// TwinCAT 3 PLC project Syn_Visu_Test
// ProgramVersion: 3.1.4026.28
// libraries:
//   Tc2_Standard, * (Beckhoff Automation GmbH)
//   Tc2_System, * (Beckhoff Automation GmbH)
//   SynConfig,newest,Syntegon Group
//   SynVisu,newest,Syntegon Group
//   TcUnit,newest,www.tcunit.org
// project tree:
//   / PlcTask.TcTTO
//   POUs/ P_TestRun.TcPOU
//   POUs/Tests/ _FB_TestBodyComponent.TcPOU, _FB_TestComponent.TcPOU, _FB_TestConfigBodyComponent.TcPOU, _FB_TestConfigComponent.TcPOU, _FB_TestConfigMachine.TcPOU, _FB_TestConfigRobot.TcPOU, _FB_TestConfigStaging.TcPOU, _FB_TestConfigTopology.TcPOU, _FB_TestConveyor.TcPOU, _FB_TestMachine.TcPOU, _FB_TestProductRegister.TcPOU, _FB_TestRobot.TcPOU, _FB_TestXtsTrack.TcPOU, _FC_TestConfigStage.TcPOU
// (motion and I/O tree: see PLC project syn_visu)
// real-time tasks:
//   TASK PlcTask: cycle T#10ms, priority 20, ADS port 350
//   TASK TestTask: cycle T#10ms, priority 21, ADS port 351

CONFIGURATION Syn_Visu_Test
    RESOURCE PLC ON TwinCAT3
        TASK PlcTask(INTERVAL := T#10ms, PRIORITY := 21);
        PROGRAM P_TestRun WITH PlcTask : P_TestRun;
    END_RESOURCE
END_CONFIGURATION

// ---- POUs/P_TestRun.TcPOU
(****************************************************************************************************<br>
© Syntegon Group.<br>
All rights reserved, also regarding any disposal, exploitation, reproduction, editing, distribution,<br>
as well as in the event of applications for industrial property rights.<br>
*****************************************************************************************************<br>
DESCRIPTION:<br>
Runs the TcUnit unit tests of the libraries Syn_Visu and Syn_Config (the installed SynVisu and SynConfig, newest<br>
versions) once after the start: every suite in POUs/Tests (_FB_TestConfig... for Syn_Config). TcUnit writes the<br>
results to the error list (ADS log) and, through TcUnit-Runner, to an xUnit file. Tests use only the libraries'<br>
public methods and their contract structures, written as the gateway writes them.<br>
****************************************************************************************************)
PROGRAM P_TestRun
VAR
	fb_TestComponent					: _FB_TestComponent;
	fb_TestConveyor						: _FB_TestConveyor;
	fb_TestProductRegister				: _FB_TestProductRegister;
	fb_TestRobot						: _FB_TestRobot;
	fb_TestXtsTrack						: _FB_TestXtsTrack;
	fb_TestBodyComponent				: _FB_TestBodyComponent;
	fb_TestMachine						: _FB_TestMachine;
	fb_TestConfigComponent				: _FB_TestConfigComponent;
	fb_TestConfigStaging				: _FB_TestConfigStaging;
	fb_TestConfigRobot					: _FB_TestConfigRobot;
	fb_TestConfigBodyComponent			: _FB_TestConfigBodyComponent;
	fb_TestConfigMachine				: _FB_TestConfigMachine;
	fb_TestConfigTopology				: _FB_TestConfigTopology;
END_VAR

TcUnit.RUN();

END_PROGRAM

// ---- POUs/Tests/_FB_TestComponent.TcPOU
(****************************************************************************************************<br>
© Syntegon Group.<br>
All rights reserved, also regarding any disposal, exploitation, reproduction, editing, distribution,<br>
as well as in the event of applications for industrial property rights.<br>
*****************************************************************************************************<br>
DESCRIPTION:<br>
TcUnit test suite of _FB_VisuComponent: registration in the manifest (m_Register, m_Id), the symbol path<br>
taken from the instance path, and the library version reported to the gateway.<br>
*****************************************************************************************************<br>
VERSION         ¦ DATE       ¦ NAME      ¦ CHANGE<br>
Syn_Visu 9.4.0  ¦ 2026-11-09 ¦ J.Willner ¦ Unit tests<br>
Syn_Visu 10.0.0 ¦ 2026-11-14 ¦ J.Willner ¦ _FC_VisuSymbolPath<br>
****************************************************************************************************)
FUNCTION_BLOCK _FB_TestComponent EXTENDS TcUnit.FB_TestSuite
VAR
	fb_PathConveyor						: _FB_VisuConveyor;	// declared here so that its instance path is known
END_VAR

m_RegisterAddsEntry();
m_RegisterIsIdempotent();
m_RegisterRejectsIdZero();
m_RegisterRejectsUsedId();
m_RegisterRejectsFullManifest();
m_RegisterSymbolPath();
m_SymbolPathFromInstancePath();
m_VersionMatchesConstant();

(****************************************************************************************************<br>
© Syntegon Group.<br>
All rights reserved, also regarding any disposal, exploitation, reproduction, editing, distribution,<br>
as well as in the event of applications for industrial property rights.<br>
*****************************************************************************************************<br>
DESCRIPTION:<br>
A new component gets a manifest entry with its id, type and name; the config version goes up by one and the<br>
manifest reports the running library's protocol and library version.<br>
****************************************************************************************************)
METHOD PRIVATE m_RegisterAddsEntry
VAR_INST
	fb_TempConveyor						: _FB_VisuConveyor;
	TempManifest						: ST_VisuManifest;
	b_TempDone							: BOOL;	// the test ran
END_VAR
TEST('RegisterAddsEntry');
IF b_TempDone THEN
	RETURN;
END_IF
b_TempDone := TRUE;

TempManifest.nProtocolVersion := 0;
AssertTrue(Condition := fb_TempConveyor.m_Register(vio_Manifest := TempManifest, vi_udn_Id := 1, vi_str_Name := 'Infeed'),
	Message := 'm_Register accepts a new id');
AssertEquals_UINT(Expected := 1, Actual := TempManifest.nCount, Message := 'one manifest entry');
AssertEquals_UDINT(Expected := 1, Actual := TempManifest.aEntries[0].nId, Message := 'entry id');
AssertTrue(Condition := TempManifest.aEntries[0].eType = E_VisuComponentType.CONVEYOR, Message := 'entry type CONVEYOR');
AssertEquals_STRING(Expected := 'Infeed', Actual := TempManifest.aEntries[0].sName, Message := 'entry name');
AssertEquals_UDINT(Expected := 2, Actual := TempManifest.nConfigVersion, Message := 'config version 1 -> 2');
AssertEquals_UINT(Expected := VISU_GlobalConst.VISU_un_PROTOCOL_VERSION, Actual := TempManifest.nProtocolVersion,
	Message := 'protocol version reported');
AssertEquals_STRING(Expected := VISU_GlobalConst.VISU_str_LIBRARY_VERSION, Actual := TempManifest.sLibraryVersion,
	Message := 'library version reported');
AssertEquals_UDINT(Expected := 1, Actual := fb_TempConveyor.m_Id(), Message := 'm_Id gives the registered id');

TEST_FINISHED();
END_METHOD

(****************************************************************************************************<br>
© Syntegon Group.<br>
All rights reserved, also regarding any disposal, exploitation, reproduction, editing, distribution,<br>
as well as in the event of applications for industrial property rights.<br>
*****************************************************************************************************<br>
DESCRIPTION:<br>
m_Register is called every cycle: registering again with the same values keeps the single entry and the<br>
config version.<br>
****************************************************************************************************)
METHOD PRIVATE m_RegisterIsIdempotent
VAR_INST
	fb_TempConveyor						: _FB_VisuConveyor;
	TempManifest						: ST_VisuManifest;
	b_TempDone							: BOOL;	// the test ran
END_VAR
TEST('RegisterIsIdempotent');
IF b_TempDone THEN
	RETURN;
END_IF
b_TempDone := TRUE;

fb_TempConveyor.m_Register(vio_Manifest := TempManifest, vi_udn_Id := 3, vi_str_Name := 'Outfeed');
AssertTrue(Condition := fb_TempConveyor.m_Register(vio_Manifest := TempManifest, vi_udn_Id := 3, vi_str_Name := 'Outfeed'),
	Message := 'the second m_Register with the same values succeeds');
AssertEquals_UINT(Expected := 1, Actual := TempManifest.nCount, Message := 'still one manifest entry');
AssertEquals_UDINT(Expected := 2, Actual := TempManifest.nConfigVersion, Message := 'config version unchanged by the second call');

TEST_FINISHED();
END_METHOD

(****************************************************************************************************<br>
© Syntegon Group.<br>
All rights reserved, also regarding any disposal, exploitation, reproduction, editing, distribution,<br>
as well as in the event of applications for industrial property rights.<br>
*****************************************************************************************************<br>
DESCRIPTION:<br>
A manifest holding VISU_un_MAX_MANIFEST_ENTRIES entries takes no further component.<br>
****************************************************************************************************)
METHOD PRIVATE m_RegisterRejectsFullManifest
VAR_INST
	fb_TempConveyor						: _FB_VisuConveyor;
	TempManifest						: ST_VisuManifest;
	b_TempDone							: BOOL;	// the test ran
END_VAR
TEST('RegisterRejectsFullManifest');
IF b_TempDone THEN
	RETURN;
END_IF
b_TempDone := TRUE;

(* Entries with id 0 never match a new id, so the manifest only counts as full. *)
TempManifest.nCount := VISU_GlobalConst_Param.VISU_un_MAX_MANIFEST_ENTRIES;
AssertFalse(Condition := fb_TempConveyor.m_Register(vio_Manifest := TempManifest, vi_udn_Id := 1, vi_str_Name := 'Infeed'),
	Message := 'full manifest refuses a new entry');
AssertEquals_UINT(Expected := VISU_GlobalConst_Param.VISU_un_MAX_MANIFEST_ENTRIES, Actual := TempManifest.nCount,
	Message := 'entry count unchanged');
AssertEquals_UDINT(Expected := 1, Actual := TempManifest.nConfigVersion, Message := 'config version unchanged');

TEST_FINISHED();
END_METHOD

(****************************************************************************************************<br>
© Syntegon Group.<br>
All rights reserved, also regarding any disposal, exploitation, reproduction, editing, distribution,<br>
as well as in the event of applications for industrial property rights.<br>
*****************************************************************************************************<br>
DESCRIPTION:<br>
Id 0 is refused without an entry, but the manifest still reports the running library's versions.<br>
****************************************************************************************************)
METHOD PRIVATE m_RegisterRejectsIdZero
VAR_INST
	fb_TempConveyor						: _FB_VisuConveyor;
	TempManifest						: ST_VisuManifest;
	b_TempDone							: BOOL;	// the test ran
END_VAR
TEST('RegisterRejectsIdZero');
IF b_TempDone THEN
	RETURN;
END_IF
b_TempDone := TRUE;

TempManifest.nProtocolVersion := 0;
AssertFalse(Condition := fb_TempConveyor.m_Register(vio_Manifest := TempManifest, vi_udn_Id := 0, vi_str_Name := 'Infeed'),
	Message := 'm_Register refuses id 0');
AssertEquals_UINT(Expected := 0, Actual := TempManifest.nCount, Message := 'no manifest entry');
AssertEquals_UDINT(Expected := 1, Actual := TempManifest.nConfigVersion, Message := 'config version unchanged');
AssertEquals_UDINT(Expected := 0, Actual := fb_TempConveyor.m_Id(), Message := 'm_Id stays 0');
AssertEquals_UINT(Expected := VISU_GlobalConst.VISU_un_PROTOCOL_VERSION, Actual := TempManifest.nProtocolVersion,
	Message := 'protocol version reported anyway');

TEST_FINISHED();
END_METHOD

(****************************************************************************************************<br>
© Syntegon Group.<br>
All rights reserved, also regarding any disposal, exploitation, reproduction, editing, distribution,<br>
as well as in the event of applications for industrial property rights.<br>
*****************************************************************************************************<br>
DESCRIPTION:<br>
An id already used by a different entry (other type or other name) is refused; the first entry stays.<br>
****************************************************************************************************)
METHOD PRIVATE m_RegisterRejectsUsedId
VAR_INST
	fb_TempConveyor						: _FB_VisuConveyor;
	fb_TempOtherConveyor				: _FB_VisuConveyor;
	fb_TempDelta						: _FB_VisuDelta;
	TempManifest						: ST_VisuManifest;
	b_TempDone							: BOOL;	// the test ran
END_VAR
TEST('RegisterRejectsUsedId');
IF b_TempDone THEN
	RETURN;
END_IF
b_TempDone := TRUE;

fb_TempConveyor.m_Register(vio_Manifest := TempManifest, vi_udn_Id := 5, vi_str_Name := 'Infeed');
AssertFalse(Condition := fb_TempDelta.m_Register(vio_Manifest := TempManifest, vi_udn_Id := 5, vi_str_Name := 'Infeed'),
	Message := 'same id, other type: refused');
AssertFalse(Condition := fb_TempOtherConveyor.m_Register(vio_Manifest := TempManifest, vi_udn_Id := 5, vi_str_Name := 'Other'),
	Message := 'same id, other name: refused');
AssertEquals_UINT(Expected := 1, Actual := TempManifest.nCount, Message := 'still one manifest entry');
AssertEquals_UDINT(Expected := 0, Actual := fb_TempDelta.m_Id(), Message := 'refused component keeps m_Id 0');
AssertEquals_UDINT(Expected := 5, Actual := fb_TempConveyor.m_Id(), Message := 'first component keeps its id');

TEST_FINISHED();
END_METHOD

(****************************************************************************************************<br>
© Syntegon Group.<br>
All rights reserved, also regarding any disposal, exploitation, reproduction, editing, distribution,<br>
as well as in the event of applications for industrial property rights.<br>
*****************************************************************************************************<br>
DESCRIPTION:<br>
The manifest entry's symbol path is the instance path without TwinCAT project and PLC project, plus<br>
'.vo_Visu': the path the gateway reads over ADS.<br>
****************************************************************************************************)
METHOD PRIVATE m_RegisterSymbolPath
VAR_INST
	TempManifest						: ST_VisuManifest;
	b_TempDone							: BOOL;	// the test ran
END_VAR
TEST('RegisterSymbolPath');
IF b_TempDone THEN
	RETURN;
END_IF
b_TempDone := TRUE;

fb_PathConveyor.m_Register(vio_Manifest := TempManifest, vi_udn_Id := 1, vi_str_Name := 'Path');
AssertEquals_STRING(Expected := 'P_TestRun.fb_TestComponent.fb_PathConveyor.vo_Visu', Actual := TempManifest.aEntries[0].sPath,
	Message := 'symbol path of vo_Visu without TwinCAT and PLC project');

TEST_FINISHED();
END_METHOD

(****************************************************************************************************<br>
© Syntegon Group.<br>
All rights reserved, also regarding any disposal, exploitation, reproduction, editing, distribution,<br>
as well as in the event of applications for industrial property rights.<br>
*****************************************************************************************************<br>
DESCRIPTION:<br>
_FC_VisuSymbolPath, the rule both manifests use: the instance path without TwinCAT project and PLC project,<br>
plus the contract structure; a path with fewer segments is kept whole.<br>
****************************************************************************************************)
METHOD PRIVATE m_SymbolPathFromInstancePath
VAR_INST
	b_TempDone							: BOOL;	// the test ran
END_VAR
TEST('SymbolPathFromInstancePath');
IF b_TempDone THEN
	RETURN;
END_IF
b_TempDone := TRUE;

AssertEquals_STRING(Expected := 'P_VisuDemoDelta.fb_Infeed1.vo_Visu',
	Actual := _FC_VisuSymbolPath(vio_str_InstancePath := 'RPP_Visu.Syn_Visu_Demo.P_VisuDemoDelta.fb_Infeed1',
		vi_str_Member := '.vo_Visu'), Message := 'TwinCAT and PLC project left out');
AssertEquals_STRING(Expected := 'P_A.fb_B.vo_Config',
	Actual := _FC_VisuSymbolPath(vio_str_InstancePath := 'Tc.Plc.P_A.fb_B', vi_str_Member := '.vo_Config'),
	Message := 'another contract structure');
AssertEquals_STRING(Expected := 'MAIN.fb_A.vo_Visu',
	Actual := _FC_VisuSymbolPath(vio_str_InstancePath := 'MAIN.fb_A', vi_str_Member := '.vo_Visu'),
	Message := 'fewer segments: kept whole');

TEST_FINISHED();
END_METHOD

(****************************************************************************************************<br>
© Syntegon Group.<br>
All rights reserved, also regarding any disposal, exploitation, reproduction, editing, distribution,<br>
as well as in the event of applications for industrial property rights.<br>
*****************************************************************************************************<br>
DESCRIPTION:<br>
_FC_GetVersionSynVisu and VISU_str_LIBRARY_VERSION name the same version: both are bumped together.<br>
****************************************************************************************************)
METHOD PRIVATE m_VersionMatchesConstant
VAR_INST
	b_TempDone							: BOOL;	// the test ran
END_VAR
VAR
	str_TempVersion						: STRING(31);	// major.minor.revision from _FC_GetVersionSynVisu
END_VAR
TEST('VersionMatchesConstant');
IF b_TempDone THEN
	RETURN;
END_IF
b_TempDone := TRUE;

str_TempVersion := CONCAT(UINT_TO_STRING(_FC_GetVersionSynVisu(vi_n_VersionElement := 1)), '.');
str_TempVersion := CONCAT(str_TempVersion, UINT_TO_STRING(_FC_GetVersionSynVisu(vi_n_VersionElement := 2)));
str_TempVersion := CONCAT(str_TempVersion, '.');
str_TempVersion := CONCAT(str_TempVersion, UINT_TO_STRING(_FC_GetVersionSynVisu(vi_n_VersionElement := 3)));
AssertEquals_STRING(Expected := VISU_GlobalConst.VISU_str_LIBRARY_VERSION, Actual := str_TempVersion,
	Message := '_FC_GetVersionSynVisu matches VISU_str_LIBRARY_VERSION');
AssertEquals_UINT(Expected := 16#FFFF, Actual := _FC_GetVersionSynVisu(vi_n_VersionElement := 4),
	Message := 'unknown version element gives 16#FFFF');

TEST_FINISHED();
END_METHOD

END_FUNCTION_BLOCK

// ---- POUs/Tests/_FB_TestConveyor.TcPOU
(****************************************************************************************************<br>
© Syntegon Group.<br>
All rights reserved, also regarding any disposal, exploitation, reproduction, editing, distribution,<br>
as well as in the event of applications for industrial property rights.<br>
*****************************************************************************************************<br>
DESCRIPTION:<br>
TcUnit test suite of _FB_VisuConveyor's config and belt position: the config version only changes when a<br>
value does, product types, the body flag, the unwrapping of a modulo belt position and the conversion between<br>
the MCS and the conveyor's coordinate system.<br>
*****************************************************************************************************<br>
VERSION         ¦ DATE       ¦ NAME      ¦ CHANGE<br>
Syn_Visu 9.4.0  ¦ 2026-11-09 ¦ J.Willner ¦ Unit tests<br>
Syn_Visu 10.0.0 ¦ 2026-11-14 ¦ J.Willner ¦ m_SetPose; m_BeltToMcs and m_McsToBelt<br>
****************************************************************************************************)
FUNCTION_BLOCK _FB_TestConveyor EXTENDS TcUnit.FB_TestSuite

m_ConfigureChangesVersionOnce();
m_SetProductTypeAddsAndUpdates();
m_SetProductTypeRejectsFullList();
m_SetBodyVisible();
m_SetModuloBeltPosition();
m_BeltAndMcsConvert();

(****************************************************************************************************<br>
© Syntegon Group.<br>
All rights reserved, also regarding any disposal, exploitation, reproduction, editing, distribution,<br>
as well as in the event of applications for industrial property rights.<br>
*****************************************************************************************************<br>
DESCRIPTION:<br>
m_BeltToMcs places a pose of the conveyor's coordinate system in the MCS as the visualisation does (the pose's<br>
rotation turns the origin shift and the position, fRz adds up), and m_McsToBelt is its inverse, also on a<br>
tilted conveyor.<br>
****************************************************************************************************)
METHOD PRIVATE m_BeltAndMcsConvert
VAR_INST
	fb_TempConveyor						: _FB_VisuConveyor;
	b_TempDone							: BOOL;	// the test ran
END_VAR
VAR
	TempPose							: ST_VisuPose;	// of the conveyor
	TempBelt							: ST_VisuPlanarPose;	// conveyor coordinate system
	TempMcs								: ST_VisuPlanarPose;
END_VAR
TEST('BeltAndMcsConvert');
IF b_TempDone THEN
	RETURN;
END_IF
b_TempDone := TRUE;


(****************************************************************************************************
A CONVEYOR TURNED BY 90 DEGREES
****************************************************************************************************)
TempPose.fX := 1000;
TempPose.fY := 500;
TempPose.fZ := 800;
TempPose.fRz := 90;
fb_TempConveyor.m_SetPose(vi_Pose := TempPose);
fb_TempConveyor.m_SetOriginShift(vi_lr_X := 100, vi_lr_Y := 0, vi_lr_Z := 0);

(* Its coordinate system lies 100 mm along the belt, i.e. along the MCS +Y. *)
TempMcs := fb_TempConveyor.m_BeltToMcs(vi_Pose := TempBelt);
AssertEquals_LREAL(Expected := 1000, Actual := TempMcs.fX, Delta := 0.001, Message := 'origin X');
AssertEquals_LREAL(Expected := 600, Actual := TempMcs.fY, Delta := 0.001, Message := 'origin Y');
AssertEquals_LREAL(Expected := 800, Actual := TempMcs.fZ, Delta := 0.001, Message := 'origin Z');
AssertEquals_LREAL(Expected := 90, Actual := TempMcs.fRz, Delta := 0.001, Message := 'origin Rz');

TempBelt.fX := 50;
TempBelt.fY := 20;
TempBelt.fZ := 10;
TempBelt.fRz := 15;
TempMcs := fb_TempConveyor.m_BeltToMcs(vi_Pose := TempBelt);
AssertEquals_LREAL(Expected := 980, Actual := TempMcs.fX, Delta := 0.001, Message := 'belt Y runs along MCS -X');
AssertEquals_LREAL(Expected := 650, Actual := TempMcs.fY, Delta := 0.001, Message := 'belt X runs along MCS +Y');
AssertEquals_LREAL(Expected := 810, Actual := TempMcs.fZ, Delta := 0.001, Message := 'Z');
AssertEquals_LREAL(Expected := 105, Actual := TempMcs.fRz, Delta := 0.001, Message := 'Rz adds up');

TempBelt := fb_TempConveyor.m_McsToBelt(vi_Pose := TempMcs);
AssertEquals_LREAL(Expected := 50, Actual := TempBelt.fX, Delta := 0.001, Message := 'back: X');
AssertEquals_LREAL(Expected := 20, Actual := TempBelt.fY, Delta := 0.001, Message := 'back: Y');
AssertEquals_LREAL(Expected := 10, Actual := TempBelt.fZ, Delta := 0.001, Message := 'back: Z');
AssertEquals_LREAL(Expected := 15, Actual := TempBelt.fRz, Delta := 0.001, Message := 'back: Rz');


(****************************************************************************************************
A TILTED CONVEYOR: THERE AND BACK
****************************************************************************************************)
TempPose.fRx := 5;
TempPose.fRy := -3;
TempPose.fRz := 30;
fb_TempConveyor.m_SetPose(vi_Pose := TempPose);
fb_TempConveyor.m_SetOriginShift(vi_lr_X := 100, vi_lr_Y := -40, vi_lr_Z := 25);
TempBelt.fX := 321;
TempBelt.fY := -45;
TempBelt.fZ := 12;
TempBelt.fRz := 7;
TempBelt := fb_TempConveyor.m_McsToBelt(vi_Pose := fb_TempConveyor.m_BeltToMcs(vi_Pose := TempBelt));
AssertEquals_LREAL(Expected := 321, Actual := TempBelt.fX, Delta := 0.001, Message := 'tilted: X');
AssertEquals_LREAL(Expected := -45, Actual := TempBelt.fY, Delta := 0.001, Message := 'tilted: Y');
AssertEquals_LREAL(Expected := 12, Actual := TempBelt.fZ, Delta := 0.001, Message := 'tilted: Z');
AssertEquals_LREAL(Expected := 7, Actual := TempBelt.fRz, Delta := 0.001, Message := 'tilted: Rz');

TEST_FINISHED();
END_METHOD

(****************************************************************************************************<br>
© Syntegon Group.<br>
All rights reserved, also regarding any disposal, exploitation, reproduction, editing, distribution,<br>
as well as in the event of applications for industrial property rights.<br>
*****************************************************************************************************<br>
DESCRIPTION:<br>
m_SetPose and m_Configure may be called every cycle: only a changed value raises the manifest's config version.<br>
****************************************************************************************************)
METHOD PRIVATE m_ConfigureChangesVersionOnce
VAR_INST
	fb_TempConveyor						: _FB_VisuConveyor;
	TempManifest						: ST_VisuManifest;
	TempPose							: ST_VisuPose;
	b_TempDone							: BOOL;	// the test ran
END_VAR
VAR
	udn_TempVersion						: UDINT;	// [-] config version after m_Register
END_VAR
TEST('ConfigureChangesVersionOnce');
IF b_TempDone THEN
	RETURN;
END_IF
b_TempDone := TRUE;

fb_TempConveyor.m_Register(vio_Manifest := TempManifest, vi_udn_Id := 1, vi_str_Name := 'Infeed');
udn_TempVersion := TempManifest.nConfigVersion;
TempPose.fX := 100;
AssertTrue(Condition := fb_TempConveyor.m_SetPose(vi_Pose := TempPose), Message := 'first m_SetPose changes the config');
AssertTrue(Condition := fb_TempConveyor.m_Configure(vi_lr_Length := 3000, vi_lr_Width := 400),
	Message := 'first m_Configure changes the config');
AssertEquals_UDINT(Expected := udn_TempVersion + 2, Actual := TempManifest.nConfigVersion,
	Message := 'config version raised once by each');
AssertFalse(Condition := fb_TempConveyor.m_SetPose(vi_Pose := TempPose), Message := 'same pose: no change');
AssertFalse(Condition := fb_TempConveyor.m_Configure(vi_lr_Length := 3000, vi_lr_Width := 400),
	Message := 'same values: no change');
AssertEquals_UDINT(Expected := udn_TempVersion + 2, Actual := TempManifest.nConfigVersion, Message := 'config version unchanged');
AssertTrue(Condition := fb_TempConveyor.m_Configure(vi_lr_Length := 3500, vi_lr_Width := 400),
	Message := 'new length changes the config');
AssertEquals_UDINT(Expected := udn_TempVersion + 3, Actual := TempManifest.nConfigVersion, Message := 'config version raised again');
AssertEquals_LREAL(Expected := 3500, Actual := fb_TempConveyor.vo_Visu.stConfig.fLength, Delta := 0.001,
	Message := 'length taken over');
AssertEquals_LREAL(Expected := 100, Actual := fb_TempConveyor.vo_Visu.stConfig.stPose.fX, Delta := 0.001,
	Message := 'pose kept by m_Configure');

TEST_FINISHED();
END_METHOD

(****************************************************************************************************<br>
© Syntegon Group.<br>
All rights reserved, also regarding any disposal, exploitation, reproduction, editing, distribution,<br>
as well as in the event of applications for industrial property rights.<br>
*****************************************************************************************************<br>
DESCRIPTION:<br>
A conveyor has a body by default; m_SetBodyVisible(FALSE) removes it once.<br>
****************************************************************************************************)
METHOD PRIVATE m_SetBodyVisible
VAR_INST
	fb_TempConveyor						: _FB_VisuConveyor;
	b_TempDone							: BOOL;	// the test ran
END_VAR
TEST('SetBodyVisible');
IF b_TempDone THEN
	RETURN;
END_IF
b_TempDone := TRUE;

AssertTrue(Condition := fb_TempConveyor.vo_Visu.stConfig.bBody, Message := 'a body by default');
AssertTrue(Condition := fb_TempConveyor.m_SetBodyVisible(vi_b_Visible := FALSE), Message := 'removing the body is a change');
AssertFalse(Condition := fb_TempConveyor.vo_Visu.stConfig.bBody, Message := 'no body');
AssertFalse(Condition := fb_TempConveyor.m_SetBodyVisible(vi_b_Visible := FALSE), Message := 'same value: no change');

TEST_FINISHED();
END_METHOD

(****************************************************************************************************<br>
© Syntegon Group.<br>
All rights reserved, also regarding any disposal, exploitation, reproduction, editing, distribution,<br>
as well as in the event of applications for industrial property rights.<br>
*****************************************************************************************************<br>
DESCRIPTION:<br>
m_SetModuloBeltPosition unwraps a modulo axis into a continuous belt position, forwards and backwards across<br>
the wrap; a reset restarts it, a period of 0 passes the position through.<br>
****************************************************************************************************)
METHOD PRIVATE m_SetModuloBeltPosition
VAR_INST
	fb_TempConveyor						: _FB_VisuConveyor;
	b_TempDone							: BOOL;	// the test ran
END_VAR
TEST('SetModuloBeltPosition');
IF b_TempDone THEN
	RETURN;
END_IF
b_TempDone := TRUE;

fb_TempConveyor.m_SetModuloBeltPosition(vi_lr_ModuloPosition := 900, vi_lr_ModuloPeriod := 1000, vi_b_Reset := FALSE);
AssertEquals_LREAL(Expected := 900, Actual := fb_TempConveyor.m_BeltPosition(), Delta := 0.001,
	Message := 'first call starts at the modulo position');
fb_TempConveyor.m_SetModuloBeltPosition(vi_lr_ModuloPosition := 100, vi_lr_ModuloPeriod := 1000, vi_b_Reset := FALSE);
AssertEquals_LREAL(Expected := 1100, Actual := fb_TempConveyor.m_BeltPosition(), Delta := 0.001,
	Message := 'forwards across the wrap');
fb_TempConveyor.m_SetModuloBeltPosition(vi_lr_ModuloPosition := 950, vi_lr_ModuloPeriod := 1000, vi_b_Reset := FALSE);
AssertEquals_LREAL(Expected := 950, Actual := fb_TempConveyor.m_BeltPosition(), Delta := 0.001,
	Message := 'backwards across the wrap');
fb_TempConveyor.m_SetModuloBeltPosition(vi_lr_ModuloPosition := 10, vi_lr_ModuloPeriod := 1000, vi_b_Reset := TRUE);
AssertEquals_LREAL(Expected := 10, Actual := fb_TempConveyor.m_BeltPosition(), Delta := 0.001,
	Message := 'reset restarts at the modulo position');
fb_TempConveyor.m_SetModuloBeltPosition(vi_lr_ModuloPosition := 123, vi_lr_ModuloPeriod := 0, vi_b_Reset := FALSE);
AssertEquals_LREAL(Expected := 123, Actual := fb_TempConveyor.m_BeltPosition(), Delta := 0.001,
	Message := 'period 0 passes the position through');

TEST_FINISHED();
END_METHOD

(****************************************************************************************************<br>
© Syntegon Group.<br>
All rights reserved, also regarding any disposal, exploitation, reproduction, editing, distribution,<br>
as well as in the event of applications for industrial property rights.<br>
*****************************************************************************************************<br>
DESCRIPTION:<br>
m_SetProductType adds a type per new id and updates the one with a known id; id 0 is refused. Setting the<br>
same values again succeeds without raising the config version.<br>
****************************************************************************************************)
METHOD PRIVATE m_SetProductTypeAddsAndUpdates
VAR_INST
	fb_TempConveyor						: _FB_VisuConveyor;
	TempManifest						: ST_VisuManifest;
	b_TempDone							: BOOL;	// the test ran
END_VAR
TEST('SetProductTypeAddsAndUpdates');
IF b_TempDone THEN
	RETURN;
END_IF
b_TempDone := TRUE;

fb_TempConveyor.m_Register(vio_Manifest := TempManifest, vi_udn_Id := 1, vi_str_Name := 'Infeed');
AssertTrue(Condition := fb_TempConveyor.m_SetProductType(vi_udn_Id := 1, vi_lr_Length := 120, vi_lr_Width := 80,
	vi_lr_Height := 40, vi_e_Shape := E_VisuProductShape.BOX, vi_lr_CornerRadius := 0), Message := 'type 1 added');
AssertTrue(Condition := fb_TempConveyor.m_SetProductType(vi_udn_Id := 2, vi_lr_Length := 66, vi_lr_Width := 66,
	vi_lr_Height := 120, vi_e_Shape := E_VisuProductShape.CYLINDER, vi_lr_CornerRadius := 0), Message := 'type 2 added');
AssertTrue(Condition := fb_TempConveyor.m_SetProductType(vi_udn_Id := 1, vi_lr_Length := 150, vi_lr_Width := 80,
	vi_lr_Height := 40, vi_e_Shape := E_VisuProductShape.ROUNDED_BOX, vi_lr_CornerRadius := 10), Message := 'type 1 updated');
AssertEquals_UINT(Expected := 2, Actual := fb_TempConveyor.vo_Visu.stConfig.nProductTypeCount, Message := 'two types');
AssertEquals_LREAL(Expected := 150, Actual := fb_TempConveyor.vo_Visu.stConfig.aProductTypes[0].fLength, Delta := 0.001,
	Message := 'type 1 length updated in place');
AssertTrue(Condition := fb_TempConveyor.vo_Visu.stConfig.aProductTypes[0].eShape = E_VisuProductShape.ROUNDED_BOX,
	Message := 'type 1 shape updated');
AssertEquals_UDINT(Expected := 5, Actual := TempManifest.nConfigVersion, Message := 'one config version per change');

AssertTrue(Condition := fb_TempConveyor.m_SetProductType(vi_udn_Id := 1, vi_lr_Length := 150, vi_lr_Width := 80,
	vi_lr_Height := 40, vi_e_Shape := E_VisuProductShape.ROUNDED_BOX, vi_lr_CornerRadius := 10),
	Message := 'same values again succeed');
AssertEquals_UDINT(Expected := 5, Actual := TempManifest.nConfigVersion, Message := 'same values: config version unchanged');

AssertFalse(Condition := fb_TempConveyor.m_SetProductType(vi_udn_Id := 0, vi_lr_Length := 10, vi_lr_Width := 10,
	vi_lr_Height := 10, vi_e_Shape := E_VisuProductShape.BOX, vi_lr_CornerRadius := 0), Message := 'id 0 refused');
AssertEquals_UINT(Expected := 2, Actual := fb_TempConveyor.vo_Visu.stConfig.nProductTypeCount, Message := 'still two types');

TEST_FINISHED();
END_METHOD

(****************************************************************************************************<br>
© Syntegon Group.<br>
All rights reserved, also regarding any disposal, exploitation, reproduction, editing, distribution,<br>
as well as in the event of applications for industrial property rights.<br>
*****************************************************************************************************<br>
DESCRIPTION:<br>
A conveyor takes VISU_un_MAX_PRODUCT_TYPES product types; a further new id is refused.<br>
****************************************************************************************************)
METHOD PRIVATE m_SetProductTypeRejectsFullList
VAR_INST
	fb_TempConveyor						: _FB_VisuConveyor;
	b_TempDone							: BOOL;	// the test ran
END_VAR
VAR
	un_TempType							: UINT;
	b_TempAllAdded						: BOOL;
END_VAR
TEST('SetProductTypeRejectsFullList');
IF b_TempDone THEN
	RETURN;
END_IF
b_TempDone := TRUE;

b_TempAllAdded := TRUE;
FOR un_TempType := 1 TO VISU_GlobalConst_Param.VISU_un_MAX_PRODUCT_TYPES DO
	b_TempAllAdded := b_TempAllAdded AND fb_TempConveyor.m_SetProductType(vi_udn_Id := UINT_TO_UDINT(un_TempType),
		vi_lr_Length := 100, vi_lr_Width := 100, vi_lr_Height := 100, vi_e_Shape := E_VisuProductShape.BOX,
		vi_lr_CornerRadius := 0);
END_FOR
AssertTrue(Condition := b_TempAllAdded, Message := 'every type up to the limit added');
AssertFalse(Condition := fb_TempConveyor.m_SetProductType(vi_udn_Id := 999, vi_lr_Length := 100, vi_lr_Width := 100,
	vi_lr_Height := 100, vi_e_Shape := E_VisuProductShape.BOX, vi_lr_CornerRadius := 0), Message := 'one more refused');
AssertEquals_UINT(Expected := VISU_GlobalConst_Param.VISU_un_MAX_PRODUCT_TYPES,
	Actual := fb_TempConveyor.vo_Visu.stConfig.nProductTypeCount, Message := 'type count at the limit');

TEST_FINISHED();
END_METHOD

END_FUNCTION_BLOCK

// ---- POUs/Tests/_FB_TestProductRegister.TcPOU
(****************************************************************************************************<br>
© Syntegon Group.<br>
All rights reserved, also regarding any disposal, exploitation, reproduction, editing, distribution,<br>
as well as in the event of applications for industrial property rights.<br>
*****************************************************************************************************<br>
DESCRIPTION:<br>
TcUnit test suite of _FB_VisuConveyor's product register: latching, the product index by id (also with a<br>
full register and after removals), product states, poses moved by the belt travel and the housekeeping of<br>
m_RemoveProductsBeyond, product marks and their names in the manifest.<br>
*****************************************************************************************************<br>
VERSION         ¦ DATE       ¦ NAME      ¦ CHANGE<br>
Syn_Visu 9.4.0  ¦ 2026-11-09 ¦ J.Willner ¦ Unit tests<br>
Syn_Visu 9.6.0  ¦ 2026-11-12 ¦ J.Willner ¦ Product marks<br>
****************************************************************************************************)
FUNCTION_BLOCK _FB_TestProductRegister EXTENDS TcUnit.FB_TestSuite

m_LatchAddsProduct();
m_LatchUsesGivenBeltPosition();
m_LatchRejectsZeroAndDuplicateId();
m_LatchFillsRegister();
m_GetProductMovesWithBelt();
m_RemoveProductKeepsOrder();
m_SetProductStateKeepsPrevious();
m_MoveProduct();
m_RemoveProductsBeyond();
m_SetProductMarkKeepsMark();
m_SetMarkNameChangesVersionOnce();

(****************************************************************************************************<br>
© Syntegon Group.<br>
All rights reserved, also regarding any disposal, exploitation, reproduction, editing, distribution,<br>
as well as in the event of applications for industrial property rights.<br>
*****************************************************************************************************<br>
DESCRIPTION:<br>
m_GetProduct gives the latch pose moved along the belt's X by the belt travel since the latch; an index out<br>
of range gives FALSE.<br>
****************************************************************************************************)
METHOD PRIVATE m_GetProductMovesWithBelt
VAR_INST
	fb_TempConveyor						: _FB_VisuConveyor;
	TempProduct							: ST_VisuProduct;
	TempPose							: ST_VisuPlanarPose;
	b_TempDone							: BOOL;	// the test ran
END_VAR
TEST('GetProductMovesWithBelt');
IF b_TempDone THEN
	RETURN;
END_IF
b_TempDone := TRUE;

fb_TempConveyor.m_SetBeltPosition(vi_lr_Position := 100);
m_Latch(vio_Conveyor := fb_TempConveyor, vi_udn_Id := 1, vi_lr_X := 50);
fb_TempConveyor.m_SetBeltPosition(vi_lr_Position := 350);
AssertTrue(Condition := fb_TempConveyor.m_GetProduct(vi_un_Index := 0, vo_Product => TempProduct, vo_Pose => TempPose),
	Message := 'index 0 exists');
AssertEquals_UDINT(Expected := 1, Actual := TempProduct.nId, Message := 'product 1');
AssertEquals_LREAL(Expected := 300, Actual := TempPose.fX, Delta := 0.001, Message := 'latch X 50 + belt travel 250');
AssertFalse(Condition := fb_TempConveyor.m_GetProduct(vi_un_Index := 1, vo_Product => TempProduct, vo_Pose => TempPose),
	Message := 'index 1 out of range');

TEST_FINISHED();
END_METHOD

(****************************************************************************************************<br>
© Syntegon Group.<br>
All rights reserved, also regarding any disposal, exploitation, reproduction, editing, distribution,<br>
as well as in the event of applications for industrial property rights.<br>
*****************************************************************************************************<br>
DESCRIPTION:<br>
Test helper: latches product vi_udn_Id as DETECTED at vi_lr_X (conveyor coordinates) and the current belt<br>
position, product type 1, no client. Result of m_LatchProduct.<br>
****************************************************************************************************)
METHOD PRIVATE m_Latch : BOOL
VAR_IN_OUT
	vio_Conveyor						: _FB_VisuConveyor;
END_VAR
VAR_INPUT
	vi_udn_Id							: UDINT;	// [-] product id
	vi_lr_X								: LREAL;	// [mm] latch pose X in the conveyor's coordinate system
END_VAR
VAR
	TempPose							: ST_VisuPlanarPose;
END_VAR
TempPose.fX := vi_lr_X;
m_Latch := vio_Conveyor.m_LatchProduct(vi_udn_Id := vi_udn_Id, vi_LatchPose := TempPose, vi_udn_ProductType := 1,
	vi_lr_LatchBeltPosition := 0, vi_b_UseLatchBeltPosition := FALSE, vi_e_State := E_VisuProductState.DETECTED,
	vi_udn_ClientId := 0);
END_METHOD

(****************************************************************************************************<br>
© Syntegon Group.<br>
All rights reserved, also regarding any disposal, exploitation, reproduction, editing, distribution,<br>
as well as in the event of applications for industrial property rights.<br>
*****************************************************************************************************<br>
DESCRIPTION:<br>
m_LatchProduct adds a valid entry with the given pose, type, state and client at the current belt position,<br>
its previous state equal to its state, no mover and no finger, and stamps the state.<br>
****************************************************************************************************)
METHOD PRIVATE m_LatchAddsProduct
VAR_INST
	fb_TempConveyor						: _FB_VisuConveyor;
	TempPose							: ST_VisuPlanarPose;
	b_TempDone							: BOOL;	// the test ran
END_VAR
TEST('LatchAddsProduct');
IF b_TempDone THEN
	RETURN;
END_IF
b_TempDone := TRUE;

fb_TempConveyor.m_SetBeltPosition(vi_lr_Position := 100);
TempPose.fX := 50;
TempPose.fY := 20;
TempPose.fRz := 90;
AssertTrue(Condition := fb_TempConveyor.m_LatchProduct(vi_udn_Id := 7, vi_LatchPose := TempPose, vi_udn_ProductType := 2,
	vi_lr_LatchBeltPosition := 0, vi_b_UseLatchBeltPosition := FALSE, vi_e_State := E_VisuProductState.DETECTED,
	vi_udn_ClientId := 60), Message := 'm_LatchProduct accepts a new id');
AssertEquals_UINT(Expected := 1, Actual := fb_TempConveyor.m_ProductCount(), Message := 'one product');
AssertEquals_UDINT(Expected := 7, Actual := fb_TempConveyor.vo_Visu.stState.aProducts[0].nId, Message := 'product id');
AssertTrue(Condition := fb_TempConveyor.vo_Visu.stState.aProducts[0].bValid, Message := 'entry valid');
AssertEquals_LREAL(Expected := 100, Actual := fb_TempConveyor.vo_Visu.stState.aProducts[0].fLatchBeltPosition, Delta := 0.001,
	Message := 'latched at the current belt position');
AssertEquals_LREAL(Expected := 20, Actual := fb_TempConveyor.vo_Visu.stState.aProducts[0].stLatchPose.fY, Delta := 0.001,
	Message := 'latch pose taken over');
AssertTrue(Condition := fb_TempConveyor.vo_Visu.stState.aProducts[0].eState = E_VisuProductState.DETECTED,
	Message := 'state DETECTED');
AssertTrue(Condition := fb_TempConveyor.vo_Visu.stState.aProducts[0].ePreviousState = E_VisuProductState.DETECTED,
	Message := 'previous state equals the state it enters in');
AssertEquals_UDINT(Expected := 60, Actual := fb_TempConveyor.vo_Visu.stState.aProducts[0].nLastClientId,
	Message := 'client that latched it');
AssertEquals_UDINT(Expected := 2, Actual := fb_TempConveyor.vo_Visu.stState.aProducts[0].nProductType, Message := 'product type');
AssertEquals_UDINT(Expected := 0, Actual := fb_TempConveyor.vo_Visu.stState.aProducts[0].nMoverId, Message := 'no mover');
AssertEquals_UDINT(Expected := 0, Actual := fb_TempConveyor.vo_Visu.stState.aProducts[0].nFingerId, Message := 'no finger');
AssertTrue(Condition := fb_TempConveyor.vo_Visu.stState.nTimestamp > 0, Message := 'state stamped with the DC time');

TEST_FINISHED();
END_METHOD

(****************************************************************************************************<br>
© Syntegon Group.<br>
All rights reserved, also regarding any disposal, exploitation, reproduction, editing, distribution,<br>
as well as in the event of applications for industrial property rights.<br>
*****************************************************************************************************<br>
DESCRIPTION:<br>
The register takes VISU_un_MAX_PRODUCTS products and refuses one more; the product index finds the first, a<br>
middle and the last one, also after a removal in the middle moved the register up.<br>
****************************************************************************************************)
METHOD PRIVATE m_LatchFillsRegister
VAR_INST
	fb_TempConveyor						: _FB_VisuConveyor;
	b_TempDone							: BOOL;	// the test ran
END_VAR
VAR
	un_TempIndex						: UINT;
	b_TempAllLatched					: BOOL;
	udn_TempMax							: UDINT;	// [-] VISU_un_MAX_PRODUCTS as an id
END_VAR
TEST('LatchFillsRegister');
IF b_TempDone THEN
	RETURN;
END_IF
b_TempDone := TRUE;

(* Ids 1000, 1001, ...: not the register indices, so a mix-up of id and index shows. *)
b_TempAllLatched := TRUE;
FOR un_TempIndex := 0 TO VISU_GlobalConst_Param.VISU_un_MAX_PRODUCTS - 1 DO
	b_TempAllLatched := b_TempAllLatched AND m_Latch(vio_Conveyor := fb_TempConveyor,
		vi_udn_Id := 1000 + UINT_TO_UDINT(un_TempIndex), vi_lr_X := 0);
END_FOR
udn_TempMax := UINT_TO_UDINT(VISU_GlobalConst_Param.VISU_un_MAX_PRODUCTS);
AssertTrue(Condition := b_TempAllLatched, Message := 'every product up to the limit latched');
AssertEquals_UINT(Expected := VISU_GlobalConst_Param.VISU_un_MAX_PRODUCTS, Actual := fb_TempConveyor.m_ProductCount(),
	Message := 'register full');
AssertFalse(Condition := m_Latch(vio_Conveyor := fb_TempConveyor, vi_udn_Id := 1, vi_lr_X := 0),
	Message := 'full register refuses one more');

AssertEquals_INT(Expected := 0, Actual := fb_TempConveyor.m_FindProduct(vi_udn_Id := 1000), Message := 'first product found');
AssertEquals_INT(Expected := 2000, Actual := fb_TempConveyor.m_FindProduct(vi_udn_Id := 3000), Message := 'middle product found');
AssertEquals_INT(Expected := UINT_TO_INT(VISU_GlobalConst_Param.VISU_un_MAX_PRODUCTS) - 1,
	Actual := fb_TempConveyor.m_FindProduct(vi_udn_Id := 1000 + udn_TempMax - 1), Message := 'last product found');
AssertEquals_INT(Expected := -1, Actual := fb_TempConveyor.m_FindProduct(vi_udn_Id := 1000 + udn_TempMax),
	Message := 'unknown id not found');

AssertTrue(Condition := fb_TempConveyor.m_RemoveProduct(vi_udn_Id := 3000), Message := 'middle product removed');
AssertEquals_INT(Expected := 2000, Actual := fb_TempConveyor.m_FindProduct(vi_udn_Id := 3001),
	Message := 'next product moved up into its place');
AssertEquals_INT(Expected := UINT_TO_INT(VISU_GlobalConst_Param.VISU_un_MAX_PRODUCTS) - 2,
	Actual := fb_TempConveyor.m_FindProduct(vi_udn_Id := 1000 + udn_TempMax - 1), Message := 'last product moved up');
AssertTrue(Condition := m_Latch(vio_Conveyor := fb_TempConveyor, vi_udn_Id := 1, vi_lr_X := 0),
	Message := 'room for one product again');

TEST_FINISHED();
END_METHOD

(****************************************************************************************************<br>
© Syntegon Group.<br>
All rights reserved, also regarding any disposal, exploitation, reproduction, editing, distribution,<br>
as well as in the event of applications for industrial property rights.<br>
*****************************************************************************************************<br>
DESCRIPTION:<br>
m_LatchProduct refuses id 0 and an id already in the register.<br>
****************************************************************************************************)
METHOD PRIVATE m_LatchRejectsZeroAndDuplicateId
VAR_INST
	fb_TempConveyor						: _FB_VisuConveyor;
	b_TempDone							: BOOL;	// the test ran
END_VAR
TEST('LatchRejectsZeroAndDuplicateId');
IF b_TempDone THEN
	RETURN;
END_IF
b_TempDone := TRUE;

AssertFalse(Condition := m_Latch(vio_Conveyor := fb_TempConveyor, vi_udn_Id := 0, vi_lr_X := 0), Message := 'id 0 refused');
AssertTrue(Condition := m_Latch(vio_Conveyor := fb_TempConveyor, vi_udn_Id := 4, vi_lr_X := 0), Message := 'id 4 latched');
AssertFalse(Condition := m_Latch(vio_Conveyor := fb_TempConveyor, vi_udn_Id := 4, vi_lr_X := 10), Message := 'id 4 again refused');
AssertEquals_UINT(Expected := 1, Actual := fb_TempConveyor.m_ProductCount(), Message := 'one product');

TEST_FINISHED();
END_METHOD

(****************************************************************************************************<br>
© Syntegon Group.<br>
All rights reserved, also regarding any disposal, exploitation, reproduction, editing, distribution,<br>
as well as in the event of applications for industrial property rights.<br>
*****************************************************************************************************<br>
DESCRIPTION:<br>
With vi_b_UseLatchBeltPosition the product is latched at the given belt position (e.g. from a touch probe),<br>
not at the current one; a robot's product enters as PLACED.<br>
****************************************************************************************************)
METHOD PRIVATE m_LatchUsesGivenBeltPosition
VAR_INST
	fb_TempConveyor						: _FB_VisuConveyor;
	TempPose							: ST_VisuPlanarPose;
	b_TempDone							: BOOL;	// the test ran
END_VAR
TEST('LatchUsesGivenBeltPosition');
IF b_TempDone THEN
	RETURN;
END_IF
b_TempDone := TRUE;

fb_TempConveyor.m_SetBeltPosition(vi_lr_Position := 100);
AssertTrue(Condition := fb_TempConveyor.m_LatchProduct(vi_udn_Id := 1, vi_LatchPose := TempPose, vi_udn_ProductType := 1,
	vi_lr_LatchBeltPosition := 80, vi_b_UseLatchBeltPosition := TRUE, vi_e_State := E_VisuProductState.PLACED,
	vi_udn_ClientId := 10), Message := 'latched');
AssertEquals_LREAL(Expected := 80, Actual := fb_TempConveyor.vo_Visu.stState.aProducts[0].fLatchBeltPosition, Delta := 0.001,
	Message := 'latched at the given belt position');
AssertTrue(Condition := fb_TempConveyor.vo_Visu.stState.aProducts[0].eState = E_VisuProductState.PLACED,
	Message := 'entered as PLACED');
AssertTrue(Condition := fb_TempConveyor.vo_Visu.stState.aProducts[0].ePreviousState = E_VisuProductState.PLACED,
	Message := 'previous state PLACED too');

TEST_FINISHED();
END_METHOD

(****************************************************************************************************<br>
© Syntegon Group.<br>
All rights reserved, also regarding any disposal, exploitation, reproduction, editing, distribution,<br>
as well as in the event of applications for industrial property rights.<br>
*****************************************************************************************************<br>
DESCRIPTION:<br>
m_MoveProduct puts a product at a new pose at the current belt position, from where the belt travel moves it<br>
on; its state stays. An unknown product gives FALSE.<br>
****************************************************************************************************)
METHOD PRIVATE m_MoveProduct
VAR_INST
	fb_TempConveyor						: _FB_VisuConveyor;
	TempProduct							: ST_VisuProduct;
	TempPose							: ST_VisuPlanarPose;
	b_TempDone							: BOOL;	// the test ran
END_VAR
TEST('MoveProduct');
IF b_TempDone THEN
	RETURN;
END_IF
b_TempDone := TRUE;

m_Latch(vio_Conveyor := fb_TempConveyor, vi_udn_Id := 1, vi_lr_X := 0);
fb_TempConveyor.m_SetProductState(vi_udn_Id := 1, vi_e_State := E_VisuProductState.ASSIGNED, vi_udn_ClientId := 10,
	vi_udn_MoverId := 0, vi_udn_FingerId := 0);
fb_TempConveyor.m_SetBeltPosition(vi_lr_Position := 200);
TempPose.fX := 500;
AssertTrue(Condition := fb_TempConveyor.m_MoveProduct(vi_udn_Id := 1, vi_Pose := TempPose), Message := 'product moved');
fb_TempConveyor.m_SetBeltPosition(vi_lr_Position := 260);
fb_TempConveyor.m_GetProduct(vi_un_Index := 0, vo_Product => TempProduct, vo_Pose => TempPose);
AssertEquals_LREAL(Expected := 560, Actual := TempPose.fX, Delta := 0.001, Message := 'new pose 500 + belt travel 60 since the move');
AssertTrue(Condition := TempProduct.eState = E_VisuProductState.ASSIGNED, Message := 'state kept');
AssertFalse(Condition := fb_TempConveyor.m_MoveProduct(vi_udn_Id := 2, vi_Pose := TempPose), Message := 'unknown product');

TEST_FINISHED();
END_METHOD

(****************************************************************************************************<br>
© Syntegon Group.<br>
All rights reserved, also regarding any disposal, exploitation, reproduction, editing, distribution,<br>
as well as in the event of applications for industrial property rights.<br>
*****************************************************************************************************<br>
DESCRIPTION:<br>
m_RemoveProduct takes a product out of the middle: the others keep their order, the freed last entry is<br>
invalid, and removing it again gives FALSE.<br>
****************************************************************************************************)
METHOD PRIVATE m_RemoveProductKeepsOrder
VAR_INST
	fb_TempConveyor						: _FB_VisuConveyor;
	b_TempDone							: BOOL;	// the test ran
END_VAR
TEST('RemoveProductKeepsOrder');
IF b_TempDone THEN
	RETURN;
END_IF
b_TempDone := TRUE;

m_Latch(vio_Conveyor := fb_TempConveyor, vi_udn_Id := 11, vi_lr_X := 0);
m_Latch(vio_Conveyor := fb_TempConveyor, vi_udn_Id := 12, vi_lr_X := 0);
m_Latch(vio_Conveyor := fb_TempConveyor, vi_udn_Id := 13, vi_lr_X := 0);
AssertTrue(Condition := fb_TempConveyor.m_RemoveProduct(vi_udn_Id := 12), Message := 'product 12 removed');
AssertEquals_UINT(Expected := 2, Actual := fb_TempConveyor.m_ProductCount(), Message := 'two products left');
AssertEquals_INT(Expected := 0, Actual := fb_TempConveyor.m_FindProduct(vi_udn_Id := 11), Message := 'product 11 stays first');
AssertEquals_INT(Expected := 1, Actual := fb_TempConveyor.m_FindProduct(vi_udn_Id := 13), Message := 'product 13 moved up');
AssertEquals_INT(Expected := -1, Actual := fb_TempConveyor.m_FindProduct(vi_udn_Id := 12), Message := 'product 12 gone');
AssertFalse(Condition := fb_TempConveyor.vo_Visu.stState.aProducts[2].bValid, Message := 'freed entry invalid');
AssertFalse(Condition := fb_TempConveyor.m_RemoveProduct(vi_udn_Id := 12), Message := 'removing it again gives FALSE');

TEST_FINISHED();
END_METHOD

(****************************************************************************************************<br>
© Syntegon Group.<br>
All rights reserved, also regarding any disposal, exploitation, reproduction, editing, distribution,<br>
as well as in the event of applications for industrial property rights.<br>
*****************************************************************************************************<br>
DESCRIPTION:<br>
m_RemoveProductsBeyond drops products that travelled beyond the given belt X, counted from the belt start<br>
(origin shift + latch X + belt travel), keeps products a robot works on wherever they are, and keeps the<br>
order and the product index of the rest.<br>
****************************************************************************************************)
METHOD PRIVATE m_RemoveProductsBeyond
VAR_INST
	fb_TempConveyor						: _FB_VisuConveyor;
	b_TempDone							: BOOL;	// the test ran
END_VAR
TEST('RemoveProductsBeyond');
IF b_TempDone THEN
	RETURN;
END_IF
b_TempDone := TRUE;

(* The conveyor's coordinate system starts 100 mm after the belt start: belt X = 100 + latch X + travel. *)
fb_TempConveyor.m_SetOriginShift(vi_lr_X := 100, vi_lr_Y := 0, vi_lr_Z := 0);
m_Latch(vio_Conveyor := fb_TempConveyor, vi_udn_Id := 1, vi_lr_X := 900);	// belt X 1000
m_Latch(vio_Conveyor := fb_TempConveyor, vi_udn_Id := 2, vi_lr_X := 950);	// belt X 1050, a robot works on it
m_Latch(vio_Conveyor := fb_TempConveyor, vi_udn_Id := 3, vi_lr_X := 200);	// belt X 300
m_Latch(vio_Conveyor := fb_TempConveyor, vi_udn_Id := 4, vi_lr_X := 960);	// belt X 1060
fb_TempConveyor.m_SetProductState(vi_udn_Id := 2, vi_e_State := E_VisuProductState.ASSIGNED, vi_udn_ClientId := 10,
	vi_udn_MoverId := 0, vi_udn_FingerId := 0);

AssertEquals_UINT(Expected := 1, Actual := fb_TempConveyor.m_RemoveProductsBeyond(vi_lr_BeltX := 1000),
	Message := 'only product 4 is beyond; product 1 on the limit stays');
AssertEquals_UINT(Expected := 3, Actual := fb_TempConveyor.m_ProductCount(), Message := 'three products left');
AssertEquals_UDINT(Expected := 1, Actual := fb_TempConveyor.vo_Visu.stState.aProducts[0].nId, Message := 'order kept: 1');
AssertEquals_UDINT(Expected := 2, Actual := fb_TempConveyor.vo_Visu.stState.aProducts[1].nId, Message := 'order kept: 2');
AssertEquals_UDINT(Expected := 3, Actual := fb_TempConveyor.vo_Visu.stState.aProducts[2].nId, Message := 'order kept: 3');
AssertFalse(Condition := fb_TempConveyor.vo_Visu.stState.aProducts[3].bValid, Message := 'freed entry invalid');

fb_TempConveyor.m_SetBeltPosition(vi_lr_Position := 100);
AssertEquals_UINT(Expected := 1, Actual := fb_TempConveyor.m_RemoveProductsBeyond(vi_lr_BeltX := 1000),
	Message := 'after 100 mm travel product 1 is beyond too; assigned product 2 stays');
AssertEquals_INT(Expected := 0, Actual := fb_TempConveyor.m_FindProduct(vi_udn_Id := 2), Message := 'product 2 moved up');
AssertEquals_INT(Expected := 1, Actual := fb_TempConveyor.m_FindProduct(vi_udn_Id := 3), Message := 'product 3 moved up');
AssertEquals_UINT(Expected := 0, Actual := fb_TempConveyor.m_RemoveProductsBeyond(vi_lr_BeltX := 1000),
	Message := 'nothing more to remove');

TEST_FINISHED();
END_METHOD

(****************************************************************************************************<br>
© Syntegon Group.<br>
All rights reserved, also regarding any disposal, exploitation, reproduction, editing, distribution,<br>
as well as in the event of applications for industrial property rights.<br>
*****************************************************************************************************<br>
DESCRIPTION:<br>
_FC_VisuSetMarkName names a mark in the manifest and bumps the config version only when the name changes;<br>
mark 0 and a mark above VISU_un_MAX_MARKS give FALSE.<br>
****************************************************************************************************)
METHOD PRIVATE m_SetMarkNameChangesVersionOnce
VAR_INST
	TempManifest						: ST_VisuManifest;
	b_TempDone							: BOOL;	// the test ran
END_VAR
TEST('SetMarkNameChangesVersionOnce');
IF b_TempDone THEN
	RETURN;
END_IF
b_TempDone := TRUE;

AssertEquals_STRING(Expected := '', Actual := TempManifest.aMarkNames[1], Message := 'unnamed at first');
AssertTrue(Condition := _FC_VisuSetMarkName(vio_Manifest := TempManifest, vi_un_Mark := 1, vi_str_Name := 'Sample'),
	Message := 'naming is a change');
AssertEquals_STRING(Expected := 'Sample', Actual := TempManifest.aMarkNames[1], Message := 'named');
AssertEquals_UDINT(Expected := 2, Actual := TempManifest.nConfigVersion, Message := 'config version bumped');
AssertFalse(Condition := _FC_VisuSetMarkName(vio_Manifest := TempManifest, vi_un_Mark := 1, vi_str_Name := 'Sample'),
	Message := 'same name: no change');
AssertEquals_UDINT(Expected := 2, Actual := TempManifest.nConfigVersion, Message := 'config version kept');

AssertFalse(Condition := _FC_VisuSetMarkName(vio_Manifest := TempManifest, vi_un_Mark := 0, vi_str_Name := 'None'),
	Message := 'mark 0 has no name');
AssertFalse(Condition := _FC_VisuSetMarkName(vio_Manifest := TempManifest,
	vi_un_Mark := VISU_GlobalConst.VISU_un_MAX_MARKS + 1, vi_str_Name := 'Too high'), Message := 'no such mark');
AssertEquals_UDINT(Expected := 2, Actual := TempManifest.nConfigVersion, Message := 'refused names change nothing');

TEST_FINISHED();
END_METHOD

(****************************************************************************************************<br>
© Syntegon Group.<br>
All rights reserved, also regarding any disposal, exploitation, reproduction, editing, distribution,<br>
as well as in the event of applications for industrial property rights.<br>
*****************************************************************************************************<br>
DESCRIPTION:<br>
A latched product is unmarked; m_SetProductMark marks it, the mark stays through m_SetProductState and<br>
m_MoveProduct, 0 removes it. A mark above VISU_un_MAX_MARKS and an unknown product give FALSE.<br>
****************************************************************************************************)
METHOD PRIVATE m_SetProductMarkKeepsMark
VAR_INST
	fb_TempConveyor						: _FB_VisuConveyor;
	TempProduct							: ST_VisuProduct;
	TempPose							: ST_VisuPlanarPose;
	b_TempDone							: BOOL;	// the test ran
END_VAR
TEST('SetProductMarkKeepsMark');
IF b_TempDone THEN
	RETURN;
END_IF
b_TempDone := TRUE;

m_Latch(vio_Conveyor := fb_TempConveyor, vi_udn_Id := 1, vi_lr_X := 0);
fb_TempConveyor.m_GetProduct(vi_un_Index := 0, vo_Product => TempProduct, vo_Pose => TempPose);
AssertEquals_UINT(Expected := 0, Actual := TempProduct.nMark, Message := 'latched unmarked');

AssertTrue(Condition := fb_TempConveyor.m_SetProductMark(vi_udn_Id := 1, vi_un_Mark := 2), Message := 'marked');
fb_TempConveyor.m_SetProductState(vi_udn_Id := 1, vi_e_State := E_VisuProductState.PICKED, vi_udn_ClientId := 10,
	vi_udn_MoverId := 0, vi_udn_FingerId := 1);
TempPose.fX := 300;
fb_TempConveyor.m_MoveProduct(vi_udn_Id := 1, vi_Pose := TempPose);
fb_TempConveyor.m_GetProduct(vi_un_Index := 0, vo_Product => TempProduct, vo_Pose => TempPose);
AssertEquals_UINT(Expected := 2, Actual := TempProduct.nMark, Message := 'mark kept through a state change and a move');

AssertFalse(Condition := fb_TempConveyor.m_SetProductMark(vi_udn_Id := 1, vi_un_Mark := VISU_GlobalConst.VISU_un_MAX_MARKS + 1),
	Message := 'no such mark');
AssertFalse(Condition := fb_TempConveyor.m_SetProductMark(vi_udn_Id := 2, vi_un_Mark := 1), Message := 'unknown product');
fb_TempConveyor.m_GetProduct(vi_un_Index := 0, vo_Product => TempProduct, vo_Pose => TempPose);
AssertEquals_UINT(Expected := 2, Actual := TempProduct.nMark, Message := 'a refused mark changes nothing');

AssertTrue(Condition := fb_TempConveyor.m_SetProductMark(vi_udn_Id := 1, vi_un_Mark := 0), Message := 'unmarked');
fb_TempConveyor.m_GetProduct(vi_un_Index := 0, vo_Product => TempProduct, vo_Pose => TempPose);
AssertEquals_UINT(Expected := 0, Actual := TempProduct.nMark, Message := 'mark removed');

TEST_FINISHED();
END_METHOD

(****************************************************************************************************<br>
© Syntegon Group.<br>
All rights reserved, also regarding any disposal, exploitation, reproduction, editing, distribution,<br>
as well as in the event of applications for industrial property rights.<br>
*****************************************************************************************************<br>
DESCRIPTION:<br>
m_SetProductState keeps the state before a change as ePreviousState (a repeated call with the same state<br>
keeps it), names the client and sets mover and finger; an unknown product gives FALSE.<br>
****************************************************************************************************)
METHOD PRIVATE m_SetProductStateKeepsPrevious
VAR_INST
	fb_TempConveyor						: _FB_VisuConveyor;
	b_TempDone							: BOOL;	// the test ran
END_VAR
TEST('SetProductStateKeepsPrevious');
IF b_TempDone THEN
	RETURN;
END_IF
b_TempDone := TRUE;

m_Latch(vio_Conveyor := fb_TempConveyor, vi_udn_Id := 1, vi_lr_X := 0);
AssertTrue(Condition := fb_TempConveyor.m_SetProductState(vi_udn_Id := 1, vi_e_State := E_VisuProductState.ASSIGNED,
	vi_udn_ClientId := 10, vi_udn_MoverId := 0, vi_udn_FingerId := 0), Message := 'assigned');
AssertTrue(Condition := fb_TempConveyor.vo_Visu.stState.aProducts[0].ePreviousState = E_VisuProductState.DETECTED,
	Message := 'previous state DETECTED');
AssertEquals_UDINT(Expected := 10, Actual := fb_TempConveyor.vo_Visu.stState.aProducts[0].nLastClientId,
	Message := 'client 10 assigned it');

fb_TempConveyor.m_SetProductState(vi_udn_Id := 1, vi_e_State := E_VisuProductState.ASSIGNED, vi_udn_ClientId := 10,
	vi_udn_MoverId := 0, vi_udn_FingerId := 0);
AssertTrue(Condition := fb_TempConveyor.vo_Visu.stState.aProducts[0].ePreviousState = E_VisuProductState.DETECTED,
	Message := 'same state again keeps the previous state');

fb_TempConveyor.m_SetProductState(vi_udn_Id := 1, vi_e_State := E_VisuProductState.PICKED, vi_udn_ClientId := 20,
	vi_udn_MoverId := 3, vi_udn_FingerId := 2);
AssertTrue(Condition := fb_TempConveyor.vo_Visu.stState.aProducts[0].eState = E_VisuProductState.PICKED,
	Message := 'state PICKED');
AssertTrue(Condition := fb_TempConveyor.vo_Visu.stState.aProducts[0].ePreviousState = E_VisuProductState.ASSIGNED,
	Message := 'previous state ASSIGNED');
AssertEquals_UDINT(Expected := 20, Actual := fb_TempConveyor.vo_Visu.stState.aProducts[0].nLastClientId,
	Message := 'client 20 picked it');
AssertEquals_UDINT(Expected := 3, Actual := fb_TempConveyor.vo_Visu.stState.aProducts[0].nMoverId, Message := 'mover 3');
AssertEquals_UDINT(Expected := 2, Actual := fb_TempConveyor.vo_Visu.stState.aProducts[0].nFingerId, Message := 'finger 2');

AssertFalse(Condition := fb_TempConveyor.m_SetProductState(vi_udn_Id := 99, vi_e_State := E_VisuProductState.REJECTED,
	vi_udn_ClientId := 70, vi_udn_MoverId := 0, vi_udn_FingerId := 0), Message := 'unknown product gives FALSE');

TEST_FINISHED();
END_METHOD

END_FUNCTION_BLOCK

// ---- POUs/Tests/_FB_TestRobot.TcPOU
(****************************************************************************************************<br>
© Syntegon Group.<br>
All rights reserved, also regarding any disposal, exploitation, reproduction, editing, distribution,<br>
as well as in the event of applications for industrial property rights.<br>
*****************************************************************************************************<br>
DESCRIPTION:<br>
TcUnit test suite of _FB_VisuZoneComponent and _FB_VisuRobot, through a Delta, a Cartesian robot and an XTS<br>
loop: zones, gripper fingers, limit area and TCP limit area, and the finger states.<br>
*****************************************************************************************************<br>
VERSION         ¦ DATE       ¦ NAME      ¦ CHANGE<br>
Syn_Visu 9.4.0  ¦ 2026-11-09 ¦ J.Willner ¦ Unit tests<br>
****************************************************************************************************)
FUNCTION_BLOCK _FB_TestRobot EXTENDS TcUnit.FB_TestSuite

m_SetZoneGrowsCount();
m_ClearZones();
m_SetFingerAndClear();
m_LimitArea();
m_TcpLimitArea();
m_XtsLoopHasNoLimitArea();
m_SetFingerState();

(****************************************************************************************************<br>
© Syntegon Group.<br>
All rights reserved, also regarding any disposal, exploitation, reproduction, editing, distribution,<br>
as well as in the event of applications for industrial property rights.<br>
*****************************************************************************************************<br>
DESCRIPTION:<br>
m_ClearZones removes every zone once (TRUE, config version raised); with no zones left it gives FALSE.<br>
****************************************************************************************************)
METHOD PRIVATE m_ClearZones
VAR_INST
	fb_TempCartesian					: _FB_VisuCartesian;
	TempManifest						: ST_VisuManifest;
	b_TempDone							: BOOL;	// the test ran
END_VAR
TEST('ClearZones');
IF b_TempDone THEN
	RETURN;
END_IF
b_TempDone := TRUE;

fb_TempCartesian.m_Register(vio_Manifest := TempManifest, vi_udn_Id := 40, vi_str_Name := 'Cartesian');
fb_TempCartesian.m_SetZone(vi_un_Zone := 1, vi_udn_ConveyorId := 7, vi_lr_Start := 1000, vi_lr_End := 2000,
	vi_lr_AllocationOffset := 0, vi_lr_CcsOffset := 1000, vi_lr_StartY := 0, vi_lr_EndY := 0);
AssertTrue(Condition := fb_TempCartesian.m_ClearZones(), Message := 'zones cleared');
AssertEquals_UINT(Expected := 0, Actual := fb_TempCartesian.vo_Visu.stConfig.nZoneCount, Message := 'no zones');
AssertEquals_UDINT(Expected := 0, Actual := fb_TempCartesian.vo_Visu.stConfig.aZones[0].nConveyorId, Message := 'zone 1 emptied');
AssertEquals_UDINT(Expected := 4, Actual := TempManifest.nConfigVersion, Message := 'config version raised by set and clear');
AssertFalse(Condition := fb_TempCartesian.m_ClearZones(), Message := 'nothing left to clear');
AssertEquals_UDINT(Expected := 4, Actual := TempManifest.nConfigVersion, Message := 'config version unchanged');

TEST_FINISHED();
END_METHOD

(****************************************************************************************************<br>
© Syntegon Group.<br>
All rights reserved, also regarding any disposal, exploitation, reproduction, editing, distribution,<br>
as well as in the event of applications for industrial property rights.<br>
*****************************************************************************************************<br>
DESCRIPTION:<br>
m_SetLimitArea activates the limit area and gives TRUE only when a value changes; m_ClearLimitArea removes<br>
it once and leaves the TCP limit area alone.<br>
****************************************************************************************************)
METHOD PRIVATE m_LimitArea
VAR_INST
	fb_TempDelta						: _FB_VisuDelta;
	TempManifest						: ST_VisuManifest;
	b_TempDone							: BOOL;	// the test ran
END_VAR
TEST('LimitArea');
IF b_TempDone THEN
	RETURN;
END_IF
b_TempDone := TRUE;

fb_TempDelta.m_Register(vio_Manifest := TempManifest, vi_udn_Id := 10, vi_str_Name := 'Delta');
AssertTrue(Condition := fb_TempDelta.m_SetLimitArea(vi_lr_XMin := -500, vi_lr_XMax := 500, vi_lr_YMin := -750,
	vi_lr_YMax := 750, vi_lr_ZMin := -1500, vi_lr_ZMax := -700), Message := 'limit area set');
AssertTrue(Condition := fb_TempDelta.vo_Visu.stConfig.stLimitArea.bActive, Message := 'limit area active');
AssertEquals_LREAL(Expected := -1500, Actual := fb_TempDelta.vo_Visu.stConfig.stLimitArea.fZMin, Delta := 0.001,
	Message := 'ZMin taken over');
AssertFalse(Condition := fb_TempDelta.vo_Visu.stConfig.stTcpLimitArea.bActive, Message := 'TCP limit area untouched');
AssertEquals_UDINT(Expected := 3, Actual := TempManifest.nConfigVersion, Message := 'config version raised');

AssertFalse(Condition := fb_TempDelta.m_SetLimitArea(vi_lr_XMin := -500, vi_lr_XMax := 500, vi_lr_YMin := -750,
	vi_lr_YMax := 750, vi_lr_ZMin := -1500, vi_lr_ZMax := -700), Message := 'same values: no change');
AssertEquals_UDINT(Expected := 3, Actual := TempManifest.nConfigVersion, Message := 'config version unchanged');

AssertTrue(Condition := fb_TempDelta.m_ClearLimitArea(), Message := 'limit area cleared');
AssertFalse(Condition := fb_TempDelta.vo_Visu.stConfig.stLimitArea.bActive, Message := 'limit area inactive');
AssertFalse(Condition := fb_TempDelta.m_ClearLimitArea(), Message := 'nothing left to clear');
AssertEquals_UDINT(Expected := 4, Actual := TempManifest.nConfigVersion, Message := 'clearing raised the config version once');

TEST_FINISHED();
END_METHOD

(****************************************************************************************************<br>
© Syntegon Group.<br>
All rights reserved, also regarding any disposal, exploitation, reproduction, editing, distribution,<br>
as well as in the event of applications for industrial property rights.<br>
*****************************************************************************************************<br>
DESCRIPTION:<br>
m_SetFinger defines a 1-based finger and grows the finger count to it; finger 0 and a finger beyond<br>
VISU_un_MAX_FINGERS are refused. m_ClearFingers removes the gripper definition once.<br>
****************************************************************************************************)
METHOD PRIVATE m_SetFingerAndClear
VAR_INST
	fb_TempXtsLoop						: _FB_VisuXtsLoop;
	b_TempDone							: BOOL;	// the test ran
END_VAR
TEST('SetFingerAndClear');
IF b_TempDone THEN
	RETURN;
END_IF
b_TempDone := TRUE;

AssertTrue(Condition := fb_TempXtsLoop.m_SetFinger(vi_un_Finger := 2, vi_lr_Diameter := 40, vi_lr_Height := 50),
	Message := 'finger 2 set');
AssertEquals_UINT(Expected := 2, Actual := fb_TempXtsLoop.vo_Visu.stConfig.nFingerCount, Message := 'finger count grows to 2');
AssertEquals_LREAL(Expected := 40, Actual := fb_TempXtsLoop.vo_Visu.stConfig.aFingers[1].fDiameter, Delta := 0.001,
	Message := 'diameter taken over');
AssertFalse(Condition := fb_TempXtsLoop.m_SetFinger(vi_un_Finger := 0, vi_lr_Diameter := 40, vi_lr_Height := 50),
	Message := 'finger 0 refused');
AssertFalse(Condition := fb_TempXtsLoop.m_SetFinger(vi_un_Finger := VISU_GlobalConst_Param.VISU_un_MAX_FINGERS + 1,
	vi_lr_Diameter := 40, vi_lr_Height := 50), Message := 'finger beyond the limit refused');

AssertTrue(Condition := fb_TempXtsLoop.m_ClearFingers(), Message := 'fingers cleared');
AssertEquals_UINT(Expected := 0, Actual := fb_TempXtsLoop.vo_Visu.stConfig.nFingerCount, Message := 'no fingers');
AssertFalse(Condition := fb_TempXtsLoop.m_ClearFingers(), Message := 'nothing left to clear');

TEST_FINISHED();
END_METHOD

(****************************************************************************************************<br>
© Syntegon Group.<br>
All rights reserved, also regarding any disposal, exploitation, reproduction, editing, distribution,<br>
as well as in the event of applications for industrial property rights.<br>
*****************************************************************************************************<br>
DESCRIPTION:<br>
A Delta's m_SetFingerState reports a 1-based finger's MCS pose and grip; finger 0 and a finger beyond<br>
VISU_un_MAX_FINGERS are refused. m_SetTcp stamps the state.<br>
****************************************************************************************************)
METHOD PRIVATE m_SetFingerState
VAR_INST
	fb_TempDelta						: _FB_VisuDelta;
	TempPose							: ST_VisuPose;
	TempTcp								: ST_VisuPosition;
	b_TempDone							: BOOL;	// the test ran
END_VAR
TEST('SetFingerState');
IF b_TempDone THEN
	RETURN;
END_IF
b_TempDone := TRUE;

TempPose.fZ := -900;
TempPose.fRz := 45;
AssertTrue(Condition := fb_TempDelta.m_SetFingerState(vi_un_Finger := 1, vi_Pose := TempPose, vi_b_Active := TRUE),
	Message := 'finger 1 reported');
AssertTrue(Condition := fb_TempDelta.vo_Visu.stState.aFingerStates[0].bActive, Message := 'finger 1 grips');
AssertEquals_LREAL(Expected := 45, Actual := fb_TempDelta.vo_Visu.stState.aFingerStates[0].stPose.fRz, Delta := 0.001,
	Message := 'finger 1 pose taken over');
AssertFalse(Condition := fb_TempDelta.m_SetFingerState(vi_un_Finger := 0, vi_Pose := TempPose, vi_b_Active := TRUE),
	Message := 'finger 0 refused');
AssertFalse(Condition := fb_TempDelta.m_SetFingerState(vi_un_Finger := VISU_GlobalConst_Param.VISU_un_MAX_FINGERS + 1,
	vi_Pose := TempPose, vi_b_Active := TRUE), Message := 'finger beyond the limit refused');

TempTcp.fZ := -1000;
fb_TempDelta.m_SetTcp(vi_ActualTcp := TempTcp, vi_SetpointTcp := TempTcp);
AssertEquals_LREAL(Expected := -1000, Actual := fb_TempDelta.vo_Visu.stState.stActualTcp.fZ, Delta := 0.001,
	Message := 'TCP taken over');
AssertTrue(Condition := fb_TempDelta.vo_Visu.stState.nTimestamp > 0, Message := 'state stamped with the DC time');

TEST_FINISHED();
END_METHOD

(****************************************************************************************************<br>
© Syntegon Group.<br>
All rights reserved, also regarding any disposal, exploitation, reproduction, editing, distribution,<br>
as well as in the event of applications for industrial property rights.<br>
*****************************************************************************************************<br>
DESCRIPTION:<br>
m_SetZone sets a 1-based zone, grows the zone count to it and raises the config version only when a value<br>
changes; zone 0, a zone beyond VISU_un_MAX_ZONES and conveyor 0 are refused.<br>
****************************************************************************************************)
METHOD PRIVATE m_SetZoneGrowsCount
VAR_INST
	fb_TempDelta						: _FB_VisuDelta;
	TempManifest						: ST_VisuManifest;
	b_TempDone							: BOOL;	// the test ran
END_VAR
TEST('SetZoneGrowsCount');
IF b_TempDone THEN
	RETURN;
END_IF
b_TempDone := TRUE;

fb_TempDelta.m_Register(vio_Manifest := TempManifest, vi_udn_Id := 10, vi_str_Name := 'Delta');
AssertTrue(Condition := fb_TempDelta.m_SetZone(vi_un_Zone := 1, vi_udn_ConveyorId := 1, vi_lr_Start := 1100, vi_lr_End := 1900,
	vi_lr_AllocationOffset := 300, vi_lr_CcsOffset := 1100, vi_lr_StartY := 0, vi_lr_EndY := 0), Message := 'zone 1 set');
AssertEquals_UINT(Expected := 1, Actual := fb_TempDelta.vo_Visu.stConfig.nZoneCount, Message := 'one zone');
AssertEquals_UDINT(Expected := 3, Actual := TempManifest.nConfigVersion, Message := 'config version raised');
AssertEquals_LREAL(Expected := 300, Actual := fb_TempDelta.vo_Visu.stConfig.aZones[0].fAllocationOffset, Delta := 0.001,
	Message := 'allocation offset taken over');

fb_TempDelta.m_SetZone(vi_un_Zone := 1, vi_udn_ConveyorId := 1, vi_lr_Start := 1100, vi_lr_End := 1900,
	vi_lr_AllocationOffset := 300, vi_lr_CcsOffset := 1100, vi_lr_StartY := 0, vi_lr_EndY := 0);
AssertEquals_UDINT(Expected := 3, Actual := TempManifest.nConfigVersion, Message := 'same zone again: config version unchanged');

AssertTrue(Condition := fb_TempDelta.m_SetZone(vi_un_Zone := 3, vi_udn_ConveyorId := 2, vi_lr_Start := 500, vi_lr_End := 900,
	vi_lr_AllocationOffset := 0, vi_lr_CcsOffset := 500, vi_lr_StartY := -100, vi_lr_EndY := 100), Message := 'zone 3 set');
AssertEquals_UINT(Expected := 3, Actual := fb_TempDelta.vo_Visu.stConfig.nZoneCount, Message := 'zone count grows to 3');
AssertEquals_LREAL(Expected := -100, Actual := fb_TempDelta.vo_Visu.stConfig.aZones[2].fStartY, Delta := 0.001,
	Message := 'lane taken over');

AssertFalse(Condition := fb_TempDelta.m_SetZone(vi_un_Zone := 0, vi_udn_ConveyorId := 1, vi_lr_Start := 0, vi_lr_End := 0,
	vi_lr_AllocationOffset := 0, vi_lr_CcsOffset := 0, vi_lr_StartY := 0, vi_lr_EndY := 0), Message := 'zone 0 refused');
AssertFalse(Condition := fb_TempDelta.m_SetZone(vi_un_Zone := VISU_GlobalConst_Param.VISU_un_MAX_ZONES + 1, vi_udn_ConveyorId := 1,
	vi_lr_Start := 0, vi_lr_End := 0, vi_lr_AllocationOffset := 0, vi_lr_CcsOffset := 0, vi_lr_StartY := 0, vi_lr_EndY := 0),
	Message := 'zone beyond the limit refused');
AssertFalse(Condition := fb_TempDelta.m_SetZone(vi_un_Zone := 2, vi_udn_ConveyorId := 0, vi_lr_Start := 0, vi_lr_End := 0,
	vi_lr_AllocationOffset := 0, vi_lr_CcsOffset := 0, vi_lr_StartY := 0, vi_lr_EndY := 0), Message := 'conveyor 0 refused');
AssertEquals_UINT(Expected := 3, Actual := fb_TempDelta.vo_Visu.stConfig.nZoneCount, Message := 'still three zones');

TEST_FINISHED();
END_METHOD

(****************************************************************************************************<br>
© Syntegon Group.<br>
All rights reserved, also regarding any disposal, exploitation, reproduction, editing, distribution,<br>
as well as in the event of applications for industrial property rights.<br>
*****************************************************************************************************<br>
DESCRIPTION:<br>
m_SetTcpLimitArea activates the TCP limit area of a Cartesian robot without touching its limit area;<br>
m_ClearTcpLimitArea removes it once.<br>
****************************************************************************************************)
METHOD PRIVATE m_TcpLimitArea
VAR_INST
	fb_TempCartesian					: _FB_VisuCartesian;
	b_TempDone							: BOOL;	// the test ran
END_VAR
TEST('TcpLimitArea');
IF b_TempDone THEN
	RETURN;
END_IF
b_TempDone := TRUE;

AssertTrue(Condition := fb_TempCartesian.m_SetTcpLimitArea(vi_lr_XMin := -60, vi_lr_XMax := 60, vi_lr_YMin := -60,
	vi_lr_YMax := 60, vi_lr_ZMin := -150, vi_lr_ZMax := 0), Message := 'TCP limit area set');
AssertTrue(Condition := fb_TempCartesian.vo_Visu.stConfig.stTcpLimitArea.bActive, Message := 'TCP limit area active');
AssertEquals_LREAL(Expected := -150, Actual := fb_TempCartesian.vo_Visu.stConfig.stTcpLimitArea.fZMin, Delta := 0.001,
	Message := 'ZMin taken over');
AssertFalse(Condition := fb_TempCartesian.vo_Visu.stConfig.stLimitArea.bActive, Message := 'limit area untouched');
AssertFalse(Condition := fb_TempCartesian.m_SetTcpLimitArea(vi_lr_XMin := -60, vi_lr_XMax := 60, vi_lr_YMin := -60,
	vi_lr_YMax := 60, vi_lr_ZMin := -150, vi_lr_ZMax := 0), Message := 'same values: no change');
AssertTrue(Condition := fb_TempCartesian.m_ClearTcpLimitArea(), Message := 'TCP limit area cleared');
AssertFalse(Condition := fb_TempCartesian.vo_Visu.stConfig.stTcpLimitArea.bActive, Message := 'TCP limit area inactive');
AssertFalse(Condition := fb_TempCartesian.m_ClearTcpLimitArea(), Message := 'nothing left to clear');

TEST_FINISHED();
END_METHOD

(****************************************************************************************************<br>
© Syntegon Group.<br>
All rights reserved, also regarding any disposal, exploitation, reproduction, editing, distribution,<br>
as well as in the event of applications for industrial property rights.<br>
*****************************************************************************************************<br>
DESCRIPTION:<br>
An XTS loop has neither a limit area nor a TCP limit area: the calls give FALSE and change no config.<br>
****************************************************************************************************)
METHOD PRIVATE m_XtsLoopHasNoLimitArea
VAR_INST
	fb_TempXtsLoop						: _FB_VisuXtsLoop;
	TempManifest						: ST_VisuManifest;
	b_TempDone							: BOOL;	// the test ran
END_VAR
TEST('XtsLoopHasNoLimitArea');
IF b_TempDone THEN
	RETURN;
END_IF
b_TempDone := TRUE;

fb_TempXtsLoop.m_Register(vio_Manifest := TempManifest, vi_udn_Id := 20, vi_str_Name := 'Fxx');
AssertFalse(Condition := fb_TempXtsLoop.m_SetLimitArea(vi_lr_XMin := -500, vi_lr_XMax := 500, vi_lr_YMin := -500,
	vi_lr_YMax := 500, vi_lr_ZMin := -500, vi_lr_ZMax := 500), Message := 'no limit area');
AssertFalse(Condition := fb_TempXtsLoop.m_SetTcpLimitArea(vi_lr_XMin := -50, vi_lr_XMax := 50, vi_lr_YMin := -50,
	vi_lr_YMax := 50, vi_lr_ZMin := -50, vi_lr_ZMax := 50), Message := 'no TCP limit area');
AssertFalse(Condition := fb_TempXtsLoop.m_ClearLimitArea(), Message := 'no limit area to clear');
AssertFalse(Condition := fb_TempXtsLoop.m_ClearTcpLimitArea(), Message := 'no TCP limit area to clear');
AssertEquals_UDINT(Expected := 2, Actual := TempManifest.nConfigVersion, Message := 'config version unchanged');

TEST_FINISHED();
END_METHOD

END_FUNCTION_BLOCK

// ---- POUs/Tests/_FB_TestXtsTrack.TcPOU
(****************************************************************************************************<br>
© Syntegon Group.<br>
All rights reserved, also regarding any disposal, exploitation, reproduction, editing, distribution,<br>
as well as in the event of applications for industrial property rights.<br>
*****************************************************************************************************<br>
DESCRIPTION:<br>
TcUnit test suite of _FB_VisuXtsTrack, _FB_VisuXtsGantry and _FB_VisuXtsLoop: track modules, the track<br>
length, module faults, the mover count and the mover entries.<br>
*****************************************************************************************************<br>
VERSION         ¦ DATE       ¦ NAME      ¦ CHANGE<br>
Syn_Visu 9.4.0  ¦ 2026-11-09 ¦ J.Willner ¦ Unit tests<br>
****************************************************************************************************)
FUNCTION_BLOCK _FB_TestXtsTrack EXTENDS TcUnit.FB_TestSuite

m_TrackLengthSumsModules();
m_SetModuleFault();
m_ClearModules();
m_MoverCount();

(****************************************************************************************************<br>
© Syntegon Group.<br>
All rights reserved, also regarding any disposal, exploitation, reproduction, editing, distribution,<br>
as well as in the event of applications for industrial property rights.<br>
*****************************************************************************************************<br>
DESCRIPTION:<br>
m_ClearModules removes the whole track once: no modules, track length 0.<br>
****************************************************************************************************)
METHOD PRIVATE m_ClearModules
VAR_INST
	fb_TempXtsGantry					: _FB_VisuXtsGantry;
	b_TempDone							: BOOL;	// the test ran
END_VAR
TEST('ClearModules');
IF b_TempDone THEN
	RETURN;
END_IF
b_TempDone := TRUE;

fb_TempXtsGantry.m_SetModule(vi_un_Module := 1, vi_e_Kind := E_VisuModuleKind.STRAIGHT,
	vi_lr_Length := VISU_GlobalConst.VISU_lr_XTS_MODULE_LENGTH);
fb_TempXtsGantry.m_SetModule(vi_un_Module := 2, vi_e_Kind := E_VisuModuleKind.STRAIGHT,
	vi_lr_Length := VISU_GlobalConst.VISU_lr_XTS_MODULE_LENGTH);
AssertTrue(Condition := fb_TempXtsGantry.m_ClearModules(), Message := 'modules cleared');
AssertEquals_UINT(Expected := 0, Actual := fb_TempXtsGantry.vo_Visu.stConfig.nModuleCount, Message := 'no modules');
AssertEquals_LREAL(Expected := 0, Actual := fb_TempXtsGantry.m_TrackLength(), Delta := 0.001, Message := 'track length 0');
AssertFalse(Condition := fb_TempXtsGantry.m_ClearModules(), Message := 'nothing left to clear');

TEST_FINISHED();
END_METHOD

(****************************************************************************************************<br>
© Syntegon Group.<br>
All rights reserved, also regarding any disposal, exploitation, reproduction, editing, distribution,<br>
as well as in the event of applications for industrial property rights.<br>
*****************************************************************************************************<br>
DESCRIPTION:<br>
m_SetMover reports a mover only inside the count set by m_SetMoverCount; lowering the count invalidates the<br>
entries beyond, a count beyond VISU_un_MAX_MOVERS is limited and gives FALSE.<br>
****************************************************************************************************)
METHOD PRIVATE m_MoverCount
VAR_INST
	fb_TempXtsGantry					: _FB_VisuXtsGantry;
	TempFingerStates					: ARRAY[0..VISU_GlobalConst_Param.VISU_un_MAX_FINGERS - 1] OF ST_VisuFingerState;
	b_TempDone							: BOOL;	// the test ran
END_VAR
TEST('MoverCount');
IF b_TempDone THEN
	RETURN;
END_IF
b_TempDone := TRUE;

AssertTrue(Condition := fb_TempXtsGantry.m_SetMoverCount(vi_un_Count := 3), Message := 'three movers');
AssertTrue(Condition := fb_TempXtsGantry.m_SetMover(vi_un_Index := 1, vi_udn_Id := 2, vi_lr_Position := 400, vi_lr_X := 120,
	vi_b_GripperActive := FALSE, vi_FingerStates := TempFingerStates, vi_b_Fault := TRUE, vi_str_FaultMessage := 'Collision'),
	Message := 'mover at index 1 reported');
AssertTrue(Condition := fb_TempXtsGantry.vo_Visu.stState.aMovers[1].bValid, Message := 'mover entry valid');
AssertEquals_LREAL(Expected := 400, Actual := fb_TempXtsGantry.vo_Visu.stState.aMovers[1].fPosition, Delta := 0.001,
	Message := 'track position taken over');
AssertTrue(Condition := fb_TempXtsGantry.vo_Visu.stState.aMovers[1].stFault.bActive, Message := 'mover fault taken over');
AssertFalse(Condition := fb_TempXtsGantry.m_SetMover(vi_un_Index := 3, vi_udn_Id := 4, vi_lr_Position := 0, vi_lr_X := 0,
	vi_b_GripperActive := FALSE, vi_FingerStates := TempFingerStates, vi_b_Fault := FALSE, vi_str_FaultMessage := ''),
	Message := 'index outside the count refused');

fb_TempXtsGantry.m_SetMoverCount(vi_un_Count := 1);
AssertFalse(Condition := fb_TempXtsGantry.vo_Visu.stState.aMovers[1].bValid, Message := 'entry beyond the new count invalid');

AssertFalse(Condition := fb_TempXtsGantry.m_SetMoverCount(vi_un_Count := VISU_GlobalConst_Param.VISU_un_MAX_MOVERS + 1),
	Message := 'count beyond the limit gives FALSE');
AssertEquals_UINT(Expected := VISU_GlobalConst_Param.VISU_un_MAX_MOVERS, Actual := fb_TempXtsGantry.vo_Visu.stState.nMoverCount,
	Message := 'count limited to VISU_un_MAX_MOVERS');

TEST_FINISHED();
END_METHOD

(****************************************************************************************************<br>
© Syntegon Group.<br>
All rights reserved, also regarding any disposal, exploitation, reproduction, editing, distribution,<br>
as well as in the event of applications for industrial property rights.<br>
*****************************************************************************************************<br>
DESCRIPTION:<br>
m_SetModuleFault sets and clears the fault of a 1-based track module in the state; module 0 is refused.<br>
****************************************************************************************************)
METHOD PRIVATE m_SetModuleFault
VAR_INST
	fb_TempXtsGantry					: _FB_VisuXtsGantry;
	b_TempDone							: BOOL;	// the test ran
END_VAR
TEST('SetModuleFault');
IF b_TempDone THEN
	RETURN;
END_IF
b_TempDone := TRUE;

AssertTrue(Condition := fb_TempXtsGantry.m_SetModuleFault(vi_un_Module := 3, vi_b_Fault := TRUE,
	vi_str_FaultMessage := 'Overtemperature'), Message := 'module 3 fault set');
AssertTrue(Condition := fb_TempXtsGantry.vo_Visu.stState.aModuleStates[2].stFault.bActive, Message := 'module 3 in a fault');
AssertEquals_STRING(Expected := 'Overtemperature', Actual := fb_TempXtsGantry.vo_Visu.stState.aModuleStates[2].stFault.sMessage,
	Message := 'fault message');
fb_TempXtsGantry.m_SetModuleFault(vi_un_Module := 3, vi_b_Fault := FALSE, vi_str_FaultMessage := '');
AssertFalse(Condition := fb_TempXtsGantry.vo_Visu.stState.aModuleStates[2].stFault.bActive, Message := 'module 3 fault cleared');
AssertFalse(Condition := fb_TempXtsGantry.m_SetModuleFault(vi_un_Module := 0, vi_b_Fault := TRUE, vi_str_FaultMessage := 'x'),
	Message := 'module 0 refused');

TEST_FINISHED();
END_METHOD

(****************************************************************************************************<br>
© Syntegon Group.<br>
All rights reserved, also regarding any disposal, exploitation, reproduction, editing, distribution,<br>
as well as in the event of applications for industrial property rights.<br>
*****************************************************************************************************<br>
DESCRIPTION:<br>
m_SetModule builds the track module by module (module 0 and one beyond VISU_un_MAX_MODULES refused), raises<br>
the config version only on a change, and m_TrackLength sums the module lengths.<br>
****************************************************************************************************)
METHOD PRIVATE m_TrackLengthSumsModules
VAR_INST
	fb_TempXtsLoop						: _FB_VisuXtsLoop;
	TempManifest						: ST_VisuManifest;
	b_TempDone							: BOOL;	// the test ran
END_VAR
VAR
	un_TempModule						: UINT;
END_VAR
TEST('TrackLengthSumsModules');
IF b_TempDone THEN
	RETURN;
END_IF
b_TempDone := TRUE;

fb_TempXtsLoop.m_Register(vio_Manifest := TempManifest, vi_udn_Id := 20, vi_str_Name := 'Fxx');
FOR un_TempModule := 1 TO 4 DO
	fb_TempXtsLoop.m_SetModule(vi_un_Module := un_TempModule, vi_e_Kind := E_VisuModuleKind.STRAIGHT,
		vi_lr_Length := VISU_GlobalConst.VISU_lr_XTS_MODULE_LENGTH);
END_FOR
AssertEquals_UINT(Expected := 4, Actual := fb_TempXtsLoop.vo_Visu.stConfig.nModuleCount, Message := 'four modules');
AssertEquals_LREAL(Expected := 1000, Actual := fb_TempXtsLoop.m_TrackLength(), Delta := 0.001, Message := '4 x 250 mm');
AssertEquals_UDINT(Expected := 6, Actual := TempManifest.nConfigVersion, Message := 'one config version per module');

fb_TempXtsLoop.m_SetModule(vi_un_Module := 2, vi_e_Kind := E_VisuModuleKind.STRAIGHT,
	vi_lr_Length := VISU_GlobalConst.VISU_lr_XTS_MODULE_LENGTH);
AssertEquals_UDINT(Expected := 6, Actual := TempManifest.nConfigVersion, Message := 'same module again: config version unchanged');

AssertTrue(Condition := fb_TempXtsLoop.m_SetModule(vi_un_Module := 2, vi_e_Kind := E_VisuModuleKind.CURVE_LEFT,
	vi_lr_Length := 125), Message := 'module 2 changed into a short curve');
AssertTrue(Condition := fb_TempXtsLoop.vo_Visu.stConfig.aModules[1].eKind = E_VisuModuleKind.CURVE_LEFT,
	Message := 'module 2 is a left curve');
AssertEquals_LREAL(Expected := 875, Actual := fb_TempXtsLoop.m_TrackLength(), Delta := 0.001, Message := 'track length 875 mm');
AssertEquals_UDINT(Expected := 7, Actual := TempManifest.nConfigVersion, Message := 'config version raised by the change');

AssertFalse(Condition := fb_TempXtsLoop.m_SetModule(vi_un_Module := 0, vi_e_Kind := E_VisuModuleKind.STRAIGHT,
	vi_lr_Length := 250), Message := 'module 0 refused');
AssertFalse(Condition := fb_TempXtsLoop.m_SetModule(vi_un_Module := VISU_GlobalConst_Param.VISU_un_MAX_MODULES + 1,
	vi_e_Kind := E_VisuModuleKind.STRAIGHT, vi_lr_Length := 250), Message := 'module beyond the limit refused');

TEST_FINISHED();
END_METHOD

END_FUNCTION_BLOCK

// ---- POUs/Tests/_FB_TestBodyComponent.TcPOU
(****************************************************************************************************<br>
© Syntegon Group.<br>
All rights reserved, also regarding any disposal, exploitation, reproduction, editing, distribution,<br>
as well as in the event of applications for industrial property rights.<br>
*****************************************************************************************************<br>
DESCRIPTION:<br>
TcUnit test suite of _FB_VisuBodyComponent through a product sensor, a vision system and a station: the bodies<br>
m_Configure describes, m_SetBody, active bodies, faults, origin shift and the state stamped by m_Register.<br>
*****************************************************************************************************<br>
VERSION         ¦ DATE       ¦ NAME      ¦ CHANGE<br>
Syn_Visu 9.4.0  ¦ 2026-11-09 ¦ J.Willner ¦ Unit tests<br>
****************************************************************************************************)
FUNCTION_BLOCK _FB_TestBodyComponent EXTENDS TcUnit.FB_TestSuite

m_SensorConfigure();
m_VisionConfigure();
m_StationBodies();
m_RegisterStampsState();

(****************************************************************************************************<br>
© Syntegon Group.<br>
All rights reserved, also regarding any disposal, exploitation, reproduction, editing, distribution,<br>
as well as in the event of applications for industrial property rights.<br>
*****************************************************************************************************<br>
DESCRIPTION:<br>
A body component may have no cyclic value of its own: its m_Register stamps the state with the DC time and<br>
enters it in the manifest with its own type.<br>
****************************************************************************************************)
METHOD PRIVATE m_RegisterStampsState
VAR_INST
	fb_TempStation						: _FB_VisuStation;
	TempManifest						: ST_VisuManifest;
	b_TempDone							: BOOL;	// the test ran
END_VAR
TEST('RegisterStampsState');
IF b_TempDone THEN
	RETURN;
END_IF
b_TempDone := TRUE;

AssertTrue(Condition := fb_TempStation.m_Register(vio_Manifest := TempManifest, vi_udn_Id := 70, vi_str_Name := 'Labeller'),
	Message := 'registered');
AssertTrue(Condition := TempManifest.aEntries[0].eType = E_VisuComponentType.STATION, Message := 'entry type STATION');
AssertTrue(Condition := fb_TempStation.vo_Visu.stState.nTimestamp > 0, Message := 'state stamped with the DC time');

TEST_FINISHED();
END_METHOD

(****************************************************************************************************<br>
© Syntegon Group.<br>
All rights reserved, also regarding any disposal, exploitation, reproduction, editing, distribution,<br>
as well as in the event of applications for industrial property rights.<br>
*****************************************************************************************************<br>
DESCRIPTION:<br>
A product sensor's m_Configure describes its head (body 1) and beam (body 2, as long as the beam), gives TRUE<br>
only on a change; m_SetPose places the head; m_SetSignal lights the beam up.<br>
****************************************************************************************************)
METHOD PRIVATE m_SensorConfigure
VAR_INST
	fb_TempSensor						: _FB_VisuSensor;
	TempManifest						: ST_VisuManifest;
	TempPose							: ST_VisuPose;
	b_TempDone							: BOOL;	// the test ran
END_VAR
TEST('SensorConfigure');
IF b_TempDone THEN
	RETURN;
END_IF
b_TempDone := TRUE;

fb_TempSensor.m_Register(vio_Manifest := TempManifest, vi_udn_Id := 61, vi_str_Name := 'Sensor');
TempPose.fX := 500;
AssertTrue(Condition := fb_TempSensor.m_SetPose(vi_Pose := TempPose), Message := 'pose set');
AssertTrue(Condition := fb_TempSensor.m_Configure(vi_lr_BeamLength := 450), Message := 'configured');
AssertEquals_UINT(Expected := 2, Actual := fb_TempSensor.vo_Visu.stConfig.nBodyCount, Message := 'head and beam');
AssertTrue(Condition := fb_TempSensor.vo_Visu.stConfig.aBodies[1].eShape = E_VisuBodyShape.CYLINDER, Message := 'beam is a cylinder');
AssertTrue(Condition := fb_TempSensor.vo_Visu.stConfig.aBodies[1].eRole = E_VisuBodyRole.BEAM, Message := 'beam role');
AssertEquals_LREAL(Expected := 450, Actual := fb_TempSensor.vo_Visu.stConfig.aBodies[1].fHeight, Delta := 0.001,
	Message := 'beam as long as configured');
AssertEquals_LREAL(Expected := 500, Actual := fb_TempSensor.vo_Visu.stConfig.stPose.fX, Delta := 0.001, Message := 'pose taken over');

AssertFalse(Condition := fb_TempSensor.m_SetPose(vi_Pose := TempPose), Message := 'same pose: no change');
AssertFalse(Condition := fb_TempSensor.m_Configure(vi_lr_BeamLength := 450), Message := 'same values: no change');

AssertTrue(Condition := fb_TempSensor.m_SetSignal(vi_b_Signal := TRUE), Message := 'signal reported');
AssertTrue(Condition := fb_TempSensor.vo_Visu.stState.aBodyStates[1].bActive, Message := 'beam lit up');
AssertFalse(Condition := fb_TempSensor.vo_Visu.stState.aBodyStates[0].bActive, Message := 'head not lit up');

TEST_FINISHED();
END_METHOD

(****************************************************************************************************<br>
© Syntegon Group.<br>
All rights reserved, also regarding any disposal, exploitation, reproduction, editing, distribution,<br>
as well as in the event of applications for industrial property rights.<br>
*****************************************************************************************************<br>
DESCRIPTION:<br>
A station describes its bodies with m_SetBody (body 0 and one beyond VISU_un_MAX_BODIES refused, the config<br>
version raised only on a change), lights one up, takes a fault and an origin shift, and m_ClearBodies<br>
removes the bodies and their active states.<br>
****************************************************************************************************)
METHOD PRIVATE m_StationBodies
VAR_INST
	fb_TempStation						: _FB_VisuStation;
	TempManifest						: ST_VisuManifest;
	TempPose							: ST_VisuPose;
	b_TempDone							: BOOL;	// the test ran
END_VAR
TEST('StationBodies');
IF b_TempDone THEN
	RETURN;
END_IF
b_TempDone := TRUE;

fb_TempStation.m_Register(vio_Manifest := TempManifest, vi_udn_Id := 70, vi_str_Name := 'Reject unit');
AssertTrue(Condition := fb_TempStation.m_SetBody(vi_un_Body := 1, vi_e_Shape := E_VisuBodyShape.BOX,
	vi_e_Role := E_VisuBodyRole.STRUCTURE, vi_Pose := TempPose, vi_lr_Length := 200, vi_lr_Width := 150, vi_lr_Height := 300,
	vi_lr_TopLength := 0, vi_lr_TopWidth := 0), Message := 'housing set');
AssertTrue(Condition := fb_TempStation.m_SetBody(vi_un_Body := 2, vi_e_Shape := E_VisuBodyShape.BOX,
	vi_e_Role := E_VisuBodyRole.STRUCTURE, vi_Pose := TempPose, vi_lr_Length := 40, vi_lr_Width := 120, vi_lr_Height := 60,
	vi_lr_TopLength := 0, vi_lr_TopWidth := 0), Message := 'pusher set');
AssertEquals_UINT(Expected := 2, Actual := fb_TempStation.vo_Visu.stConfig.nBodyCount, Message := 'two bodies');
AssertEquals_UDINT(Expected := 4, Actual := TempManifest.nConfigVersion, Message := 'one config version per body');
fb_TempStation.m_SetBody(vi_un_Body := 2, vi_e_Shape := E_VisuBodyShape.BOX, vi_e_Role := E_VisuBodyRole.STRUCTURE,
	vi_Pose := TempPose, vi_lr_Length := 40, vi_lr_Width := 120, vi_lr_Height := 60, vi_lr_TopLength := 0, vi_lr_TopWidth := 0);
AssertEquals_UDINT(Expected := 4, Actual := TempManifest.nConfigVersion, Message := 'same body again: config version unchanged');
AssertFalse(Condition := fb_TempStation.m_SetBody(vi_un_Body := 0, vi_e_Shape := E_VisuBodyShape.BOX,
	vi_e_Role := E_VisuBodyRole.STRUCTURE, vi_Pose := TempPose, vi_lr_Length := 1, vi_lr_Width := 1, vi_lr_Height := 1,
	vi_lr_TopLength := 0, vi_lr_TopWidth := 0), Message := 'body 0 refused');
AssertFalse(Condition := fb_TempStation.m_SetBody(vi_un_Body := VISU_GlobalConst_Param.VISU_un_MAX_BODIES + 1,
	vi_e_Shape := E_VisuBodyShape.BOX, vi_e_Role := E_VisuBodyRole.STRUCTURE, vi_Pose := TempPose, vi_lr_Length := 1,
	vi_lr_Width := 1, vi_lr_Height := 1, vi_lr_TopLength := 0, vi_lr_TopWidth := 0), Message := 'body beyond the limit refused');

AssertTrue(Condition := fb_TempStation.m_SetBodyActive(vi_un_Body := 2, vi_b_Active := TRUE), Message := 'pusher active');
AssertTrue(Condition := fb_TempStation.vo_Visu.stState.aBodyStates[1].bActive, Message := 'pusher lit up');

AssertTrue(Condition := fb_TempStation.m_SetFault(vi_b_Active := TRUE, vi_str_Message := 'Air pressure'), Message := 'fault set');
AssertTrue(Condition := fb_TempStation.vo_Visu.stState.stFault.bActive, Message := 'station in a fault');
AssertEquals_STRING(Expected := 'Air pressure', Actual := fb_TempStation.vo_Visu.stState.stFault.sMessage, Message := 'fault message');

AssertTrue(Condition := fb_TempStation.m_SetOriginShift(vi_lr_X := 100, vi_lr_Y := 0, vi_lr_Z := 0), Message := 'origin shifted');
AssertFalse(Condition := fb_TempStation.m_SetOriginShift(vi_lr_X := 100, vi_lr_Y := 0, vi_lr_Z := 0),
	Message := 'same origin shift: no change');

AssertTrue(Condition := fb_TempStation.m_ClearBodies(), Message := 'bodies cleared');
AssertEquals_UINT(Expected := 0, Actual := fb_TempStation.vo_Visu.stConfig.nBodyCount, Message := 'no bodies');
AssertFalse(Condition := fb_TempStation.vo_Visu.stState.aBodyStates[1].bActive, Message := 'active state cleared too');

TEST_FINISHED();
END_METHOD

